Universal Robots URScript: test_4.script

def Machining2():
  # Default parameters:
  global speed_ms = 0.3
  global speed_rads = 0.75
  global accel_mss = 3
  global accel_radss = 1.2
  global blend_radius_m = 0.001

  # Add subprograms here
  # Start of main program
  # Program generated by RoboDK v5.6.5 for UR10e on 02/02/2024 11:53:03
  # Using nominal kinematics.
  blend_radius_m = 0.002
  speed_ms = 1.000
  # set_reference(p[0.335000, -0.152000, -0.013000, 0.000000, 0.000000, 0.000000])
  set_tcp(p[0.000000, 0.000000, 0.252000, 0.000000, 0.000000, 0.000000])
  # Show Tool
  movej([0.067194, -1.005485, -2.507684, -1.199220, 1.570796, 1.637990],accel_radss,speed_rads,0,blend_radius_m)
  movel([0.067194, -1.005485, -2.507684, -1.199220, 1.570796, 1.637990],accel_mss,speed_ms,0,blend_radius_m)
  # Splitting Linear movement in 6 (instruction 7: MoveL 3)
  movel([0.067194, -1.023371, -2.532341, -1.156677, 1.570796, 1.637990],accel_mss,speed_ms,0,blend_radius_m)
  movel([0.067194, -1.043822, -2.556463, -1.112104, 1.570796, 1.637990],accel_mss,speed_ms,0,blend_radius_m)
  movel([0.067194, -1.067076, -2.580006, -1.065307, 1.570796, 1.637990],accel_mss,speed_ms,0,blend_radius_m)
  movel([0.067194, -1.093389, -2.602916, -1.016084, 1.570796, 1.637990],accel_mss,speed_ms,0,blend_radius_m)
  movel([0.067194, -1.123035, -2.625130, -0.964224, 1.570796, 1.637990],accel_mss,speed_ms,0,blend_radius_m)
  movel([0.067194, -1.156300, -2.646577, -0.909512, 1.570796, 1.637990],accel_mss,speed_ms,0,blend_radius_m)
  movel([0.067194, -1.156300, -2.646577, -0.909512, 1.570796, 1.637990],accel_mss,speed_ms,0,blend_radius_m)
  speed_ms = 1.000
  movel([0.067194, -1.156300, -2.646577, -0.909512, 1.570796, 1.637990],accel_mss,speed_ms,0,blend_radius_m)
  movel([0.067194, -1.156300, -2.646577, -0.909512, 1.570796, 1.637990],accel_mss,speed_ms,0,blend_radius_m)
  movel([0.067194, -1.156300, -2.646577, -0.909512, 1.570796, 1.637990],accel_mss,speed_ms,0,blend_radius_m)
  speed_ms = 0.005
  # Splitting Linear movement in 2 (instruction 14: MoveL 8)
  movel([0.067194, -1.135891, -2.633806, -0.942693, 1.570796, 1.637990],accel_mss,speed_ms,0,blend_radius_m)
  movel([0.067194, -1.116825, -2.620746, -0.974817, 1.570796, 1.637990],accel_mss,speed_ms,0,blend_radius_m)
  speed_ms = 1.000
  # Splitting Linear movement in 2 (instruction 16: MoveL 9)
  movel([0.067194, -1.135891, -2.633806, -0.942693, 1.570796, 1.637990],accel_mss,speed_ms,0,blend_radius_m)
  movel([0.067194, -1.156300, -2.646577, -0.909512, 1.570796, 1.637990],accel_mss,speed_ms,0,blend_radius_m)
  speed_ms = 0.040
  movel([0.067194, -1.156300, -2.646577, -0.909512, 1.570796, 1.637990],accel_mss,speed_ms,0,blend_radius_m)
  speed_ms = 1.000
  movel([0.067194, -1.156300, -2.646577, -0.909512, 1.570796, 1.637990],accel_mss,speed_ms,0,blend_radius_m)
  # Splitting Linear movement in 8 (instruction 21: MoveL 12)
  movel([0.093765, -1.178967, -2.636050, -0.897372, 1.570796, 1.664562],accel_mss,speed_ms,0,blend_radius_m)
  movel([0.118639, -1.202315, -2.624642, -0.885432, 1.570796, 1.689436],accel_mss,speed_ms,0,blend_radius_m)
  movel([0.141916, -1.226161, -2.612379, -0.873849, 1.570796, 1.712712],accel_mss,speed_ms,0,blend_radius_m)
  movel([0.163698, -1.250347, -2.599285, -0.862758, 1.570796, 1.734494],accel_mss,speed_ms,0,blend_radius_m)
  movel([0.184083, -1.274733, -2.585389, -0.852267, 1.570796, 1.754880],accel_mss,speed_ms,0,blend_radius_m)
  movel([0.203170, -1.299204, -2.570720, -0.842465, 1.570796, 1.773967],accel_mss,speed_ms,0,blend_radius_m)
  movel([0.221051, -1.323665, -2.555309, -0.833415, 1.570796, 1.791848],accel_mss,speed_ms,0,blend_radius_m)
  movel([0.237813, -1.348037, -2.539186, -0.825166, 1.570796, 1.808610],accel_mss,speed_ms,0,blend_radius_m)
  speed_ms = 0.005
  movel([0.237813, -1.389023, -2.559646, -0.763720, 1.570796, 1.808610],accel_mss,speed_ms,0,blend_radius_m)
  speed_ms = 0.025
  movel([0.235045, -1.393576, -2.556354, -0.762459, 1.570796, 1.805842],accel_mss,speed_ms,0,blend_radius_m)
  movel([0.233553, -1.395826, -2.554716, -0.761847, 1.570796, 1.804349],accel_mss,speed_ms,0,blend_radius_m)
  movel([0.231969, -1.398040, -2.553098, -0.761252, 1.570796, 1.802766],accel_mss,speed_ms,0,blend_radius_m)
  movel([0.230284, -1.400201, -2.551510, -0.760677, 1.570796, 1.801081],accel_mss,speed_ms,0,blend_radius_m)
  movel([0.228485, -1.402296, -2.549965, -0.760127, 1.570796, 1.799282],accel_mss,speed_ms,0,blend_radius_m)
  movel([0.226558, -1.404312, -2.548473, -0.759604, 1.570796, 1.797355],accel_mss,speed_ms,0,blend_radius_m)
  movel([0.224490, -1.406231, -2.547046, -0.759112, 1.570796, 1.795286],accel_mss,speed_ms,0,blend_radius_m)
  movel([0.225289, -1.405338, -2.547711, -0.759341, 1.570796, 1.796085],accel_mss,speed_ms,0,blend_radius_m)
  movel([0.226090, -1.404119, -2.548616, -0.759654, 1.570796, 1.796886],accel_mss,speed_ms,0,blend_radius_m)
  movel([0.226657, -1.402885, -2.549530, -0.759974, 1.570796, 1.797453],accel_mss,speed_ms,0,blend_radius_m)
  movel([0.226775, -1.402364, -2.549915, -0.760110, 1.570796, 1.797572],accel_mss,speed_ms,0,blend_radius_m)
  movel([0.226747, -1.401956, -2.550216, -0.760216, 1.570796, 1.797543],accel_mss,speed_ms,0,blend_radius_m)
  movel([0.226540, -1.401693, -2.550411, -0.760285, 1.570796, 1.797336],accel_mss,speed_ms,0,blend_radius_m)
  movel([0.226190, -1.401646, -2.550445, -0.760297, 1.570796, 1.796986],accel_mss,speed_ms,0,blend_radius_m)
  movel([0.225721, -1.401788, -2.550341, -0.760260, 1.570796, 1.796518],accel_mss,speed_ms,0,blend_radius_m)
  movel([0.225147, -1.402096, -2.550113, -0.760180, 1.570796, 1.795944],accel_mss,speed_ms,0,blend_radius_m)
  movel([0.223775, -1.403102, -2.549370, -0.759918, 1.570796, 1.794571],accel_mss,speed_ms,0,blend_radius_m)
  movel([0.222231, -1.404457, -2.548365, -0.759567, 1.570796, 1.793027],accel_mss,speed_ms,0,blend_radius_m)
  movel([0.219245, -1.407409, -2.546167, -0.758812, 1.570796, 1.790041],accel_mss,speed_ms,0,blend_radius_m)
  movel([0.217410, -1.409332, -2.544729, -0.758328, 1.570796, 1.788207],accel_mss,speed_ms,0,blend_radius_m)
  movel([0.214705, -1.411968, -2.542749, -0.757672, 1.570796, 1.785501],accel_mss,speed_ms,0,blend_radius_m)
  movel([0.213250, -1.413159, -2.541851, -0.757379, 1.570796, 1.784046],accel_mss,speed_ms,0,blend_radius_m)
  movel([0.211689, -1.414182, -2.541078, -0.757129, 1.570796, 1.782486],accel_mss,speed_ms,0,blend_radius_m)
  movel([0.212040, -1.413816, -2.541354, -0.757218, 1.570796, 1.782836],accel_mss,speed_ms,0,blend_radius_m)
  movel([0.212351, -1.413193, -2.541825, -0.757371, 1.570796, 1.783147],accel_mss,speed_ms,0,blend_radius_m)
  movel([0.212822, -1.411511, -2.543093, -0.757785, 1.570796, 1.783618],accel_mss,speed_ms,0,blend_radius_m)
  movel([0.213027, -1.409824, -2.544360, -0.758204, 1.570796, 1.783823],accel_mss,speed_ms,0,blend_radius_m)
  movel([0.213004, -1.409193, -2.544834, -0.758363, 1.570796, 1.783800],accel_mss,speed_ms,0,blend_radius_m)
  movel([0.212886, -1.408822, -2.545111, -0.758456, 1.570796, 1.783683],accel_mss,speed_ms,0,blend_radius_m)
  movel([0.212415, -1.408436, -2.545400, -0.758553, 1.570796, 1.783211],accel_mss,speed_ms,0,blend_radius_m)
  movel([0.211885, -1.408340, -2.545472, -0.758577, 1.570796, 1.782681],accel_mss,speed_ms,0,blend_radius_m)
  movel([0.211310, -1.408476, -2.545370, -0.758543, 1.570796, 1.782107],accel_mss,speed_ms,0,blend_radius_m)
  movel([0.210707, -1.408794, -2.545132, -0.758463, 1.570796, 1.781503],accel_mss,speed_ms,0,blend_radius_m)
  movel([0.209488, -1.409732, -2.544429, -0.758227, 1.570796, 1.780285],accel_mss,speed_ms,0,blend_radius_m)
  movel([0.208361, -1.410705, -2.543699, -0.757985, 1.570796, 1.779157],accel_mss,speed_ms,0,blend_radius_m)
  movel([0.206539, -1.412115, -2.542638, -0.757636, 1.570796, 1.777335],accel_mss,speed_ms,0,blend_radius_m)
  movel([0.204719, -1.413331, -2.541721, -0.757337, 1.570796, 1.775515],accel_mss,speed_ms,0,blend_radius_m)
  movel([0.202815, -1.414308, -2.540982, -0.757099, 1.570796, 1.773611],accel_mss,speed_ms,0,blend_radius_m)
  movel([0.200751, -1.414992, -2.540465, -0.756933, 1.570796, 1.771548],accel_mss,speed_ms,0,blend_radius_m)
  movel([0.202050, -1.413855, -2.541325, -0.757209, 1.570796, 1.772846],accel_mss,speed_ms,0,blend_radius_m)
  movel([0.203160, -1.412607, -2.542267, -0.757515, 1.570796, 1.773956],accel_mss,speed_ms,0,blend_radius_m)
  movel([0.203562, -1.411917, -2.542787, -0.757685, 1.570796, 1.774359],accel_mss,speed_ms,0,blend_radius_m)
  movel([0.203796, -1.411225, -2.543308, -0.757856, 1.570796, 1.774592],accel_mss,speed_ms,0,blend_radius_m)
  movel([0.203827, -1.410587, -2.543788, -0.758014, 1.570796, 1.774624],accel_mss,speed_ms,0,blend_radius_m)
  movel([0.203610, -1.410065, -2.544180, -0.758144, 1.570796, 1.774406],accel_mss,speed_ms,0,blend_radius_m)
  movel([0.203000, -1.409678, -2.544470, -0.758241, 1.570796, 1.773797],accel_mss,speed_ms,0,blend_radius_m)
  movel([0.202157, -1.409585, -2.544540, -0.758264, 1.570796, 1.772954],accel_mss,speed_ms,0,blend_radius_m)
  movel([0.201181, -1.409700, -2.544453, -0.758235, 1.570796, 1.771977],accel_mss,speed_ms,0,blend_radius_m)
  movel([0.200179, -1.409929, -2.544282, -0.758178, 1.570796, 1.770975],accel_mss,speed_ms,0,blend_radius_m)
  speed_ms = 0.005
  movel([0.200179, -1.401572, -2.540395, -0.770422, 1.570796, 1.770975],accel_mss,speed_ms,0,blend_radius_m)
  speed_ms = 0.040
  movel([0.198845, -1.420778, -2.525900, -0.765711, 1.570796, 1.769641],accel_mss,speed_ms,0,blend_radius_m)
  speed_ms = 0.005
  movel([0.198845, -1.428998, -2.529707, -0.753685, 1.570796, 1.769641],accel_mss,speed_ms,0,blend_radius_m)
  speed_ms = 0.025
  movel([0.199509, -1.427856, -2.530594, -0.753939, 1.570796, 1.770306],accel_mss,speed_ms,0,blend_radius_m)
  movel([0.200309, -1.426742, -2.531459, -0.754188, 1.570796, 1.771105],accel_mss,speed_ms,0,blend_radius_m)
  movel([0.201225, -1.425672, -2.532287, -0.754429, 1.570796, 1.772021],accel_mss,speed_ms,0,blend_radius_m)
  movel([0.202246, -1.424659, -2.533070, -0.754660, 1.570796, 1.773042],accel_mss,speed_ms,0,blend_radius_m)
  movel([0.203354, -1.423716, -2.533798, -0.754875, 1.570796, 1.774151],accel_mss,speed_ms,0,blend_radius_m)
  movel([0.204537, -1.422860, -2.534457, -0.755072, 1.570796, 1.775333],accel_mss,speed_ms,0,blend_radius_m)
  movel([0.205775, -1.422105, -2.535038, -0.755247, 1.570796, 1.776572],accel_mss,speed_ms,0,blend_radius_m)
  movel([0.207059, -1.421462, -2.535531, -0.755396, 1.570796, 1.777855],accel_mss,speed_ms,0,blend_radius_m)
  movel([0.208994, -1.420727, -2.536094, -0.755567, 1.570796, 1.779790],accel_mss,speed_ms,0,blend_radius_m)
  movel([0.210833, -1.420284, -2.536434, -0.755671, 1.570796, 1.781629],accel_mss,speed_ms,0,blend_radius_m)
  movel([0.212575, -1.420109, -2.536568, -0.755712, 1.570796, 1.783371],accel_mss,speed_ms,0,blend_radius_m)
  movel([0.214215, -1.420179, -2.536514, -0.755696, 1.570796, 1.785012],accel_mss,speed_ms,0,blend_radius_m)
  movel([0.215754, -1.420471, -2.536291, -0.755627, 1.570796, 1.786550],accel_mss,speed_ms,0,blend_radius_m)
  movel([0.217191, -1.420963, -2.535914, -0.755512, 1.570796, 1.787988],accel_mss,speed_ms,0,blend_radius_m)
  movel([0.218522, -1.421632, -2.535400, -0.755356, 1.570796, 1.789319],accel_mss,speed_ms,0,blend_radius_m)
  movel([0.219749, -1.422454, -2.534769, -0.755166, 1.570796, 1.790545],accel_mss,speed_ms,0,blend_radius_m)
  movel([0.220869, -1.423406, -2.534037, -0.754946, 1.570796, 1.791665],accel_mss,speed_ms,0,blend_radius_m)
  movel([0.221883, -1.424465, -2.533220, -0.754704, 1.570796, 1.792680],accel_mss,speed_ms,0,blend_radius_m)
  movel([0.223597, -1.426808, -2.531407, -0.754173, 1.570796, 1.794393],accel_mss,speed_ms,0,blend_radius_m)
  movel([0.224891, -1.429295, -2.529475, -0.753619, 1.570796, 1.795688],accel_mss,speed_ms,0,blend_radius_m)
  movel([0.225764, -1.431748, -2.527560, -0.753082, 1.570796, 1.796561],accel_mss,speed_ms,0,blend_radius_m)
  movel([0.226370, -1.434419, -2.525463, -0.752506, 1.570796, 1.797167],accel_mss,speed_ms,0,blend_radius_m)
  movel([0.226742, -1.437185, -2.523282, -0.751922, 1.570796, 1.797539],accel_mss,speed_ms,0,blend_radius_m)
  movel([0.226909, -1.440026, -2.521029, -0.751334, 1.570796, 1.797705],accel_mss,speed_ms,0,blend_radius_m)
  movel([0.226896, -1.442925, -2.518717, -0.750747, 1.570796, 1.797692],accel_mss,speed_ms,0,blend_radius_m)
  movel([0.226731, -1.445864, -2.516361, -0.750164, 1.570796, 1.797527],accel_mss,speed_ms,0,blend_radius_m)
  movel([0.226444, -1.448825, -2.513973, -0.749591, 1.570796, 1.797240],accel_mss,speed_ms,0,blend_radius_m)
  movel([0.225607, -1.454748, -2.509158, -0.748483, 1.570796, 1.796403],accel_mss,speed_ms,0,blend_radius_m)
  movel([0.224989, -1.458871, -2.505774, -0.747744, 1.570796, 1.795785],accel_mss,speed_ms,0,blend_radius_m)
  movel([0.224859, -1.460871, -2.504123, -0.747395, 1.570796, 1.795655],accel_mss,speed_ms,0,blend_radius_m)
  movel([0.224966, -1.462787, -2.502536, -0.747066, 1.570796, 1.795762],accel_mss,speed_ms,0,blend_radius_m)
  movel([0.225466, -1.465173, -2.500551, -0.746665, 1.570796, 1.796262],accel_mss,speed_ms,0,blend_radius_m)
  movel([0.225968, -1.467564, -2.498554, -0.746271, 1.570796, 1.796765],accel_mss,speed_ms,0,blend_radius_m)
  movel([0.226065, -1.468777, -2.497537, -0.746075, 1.570796, 1.796861],accel_mss,speed_ms,0,blend_radius_m)
  movel([0.225974, -1.470011, -2.496500, -0.745878, 1.570796, 1.796771],accel_mss,speed_ms,0,blend_radius_m)
  movel([0.225636, -1.471270, -2.495440, -0.745679, 1.570796, 1.796433],accel_mss,speed_ms,0,blend_radius_m)
  movel([0.224991, -1.472564, -2.494348, -0.745477, 1.570796, 1.795787],accel_mss,speed_ms,0,blend_radius_m)
  movel([0.226901, -1.469422, -2.496996, -0.745972, 1.570796, 1.797697],accel_mss,speed_ms,0,blend_radius_m)
  movel([0.228644, -1.466259, -2.499645, -0.746485, 1.570796, 1.799440],accel_mss,speed_ms,0,blend_radius_m)
  movel([0.231835, -1.459849, -2.504967, -0.747573, 1.570796, 1.802632],accel_mss,speed_ms,0,blend_radius_m)
  movel([0.233501, -1.456244, -2.507933, -0.748212, 1.570796, 1.804297],accel_mss,speed_ms,0,blend_radius_m)
  movel([0.235068, -1.452620, -2.510894, -0.748875, 1.570796, 1.805865],accel_mss,speed_ms,0,blend_radius_m)
  movel([0.237984, -1.445308, -2.516808, -0.750274, 1.570796, 1.808780],accel_mss,speed_ms,0,blend_radius_m)
  movel([0.240604, -1.438082, -2.522572, -0.751735, 1.570796, 1.811400],accel_mss,speed_ms,0,blend_radius_m)
  movel([0.241738, -1.434441, -2.525447, -0.752502, 1.570796, 1.812534],accel_mss,speed_ms,0,blend_radius_m)
  movel([0.242662, -1.430833, -2.528275, -0.753281, 1.570796, 1.813459],accel_mss,speed_ms,0,blend_radius_m)
  movel([0.243176, -1.428019, -2.530468, -0.753902, 1.570796, 1.813972],accel_mss,speed_ms,0,blend_radius_m)
  movel([0.243556, -1.425209, -2.532645, -0.754534, 1.570796, 1.814353],accel_mss,speed_ms,0,blend_radius_m)
  movel([0.243953, -1.422370, -2.534833, -0.755185, 1.570796, 1.814749],accel_mss,speed_ms,0,blend_radius_m)
  movel([0.244515, -1.419469, -2.537057, -0.755863, 1.570796, 1.815311],accel_mss,speed_ms,0,blend_radius_m)
  movel([0.244763, -1.418683, -2.537657, -0.756048, 1.570796, 1.815560],accel_mss,speed_ms,0,blend_radius_m)
  movel([0.245167, -1.417894, -2.538259, -0.756236, 1.570796, 1.815963],accel_mss,speed_ms,0,blend_radius_m)
  movel([0.245733, -1.417238, -2.538759, -0.756392, 1.570796, 1.816529],accel_mss,speed_ms,0,blend_radius_m)
  movel([0.246084, -1.417001, -2.538939, -0.756449, 1.570796, 1.816880],accel_mss,speed_ms,0,blend_radius_m)
  movel([0.246482, -1.416844, -2.539058, -0.756486, 1.570796, 1.817278],accel_mss,speed_ms,0,blend_radius_m)
  movel([0.247021, -1.416802, -2.539091, -0.756496, 1.570796, 1.817817],accel_mss,speed_ms,0,blend_radius_m)
  movel([0.247506, -1.416887, -2.539026, -0.756476, 1.570796, 1.818302],accel_mss,speed_ms,0,blend_radius_m)
  movel([0.249997, -1.417659, -2.538438, -0.756291, 1.570796, 1.820793],accel_mss,speed_ms,0,blend_radius_m)
  movel([0.252171, -1.418695, -2.537648, -0.756045, 1.570796, 1.822967],accel_mss,speed_ms,0,blend_radius_m)
  movel([0.254051, -1.419966, -2.536677, -0.755746, 1.570796, 1.824848],accel_mss,speed_ms,0,blend_radius_m)
  movel([0.255662, -1.421454, -2.535537, -0.755398, 1.570796, 1.826458],accel_mss,speed_ms,0,blend_radius_m)
  movel([0.257025, -1.423131, -2.534248, -0.755010, 1.570796, 1.827822],accel_mss,speed_ms,0,blend_radius_m)
  movel([0.258167, -1.424975, -2.532827, -0.754588, 1.570796, 1.828963],accel_mss,speed_ms,0,blend_radius_m)
  movel([0.259109, -1.426961, -2.531289, -0.754139, 1.570796, 1.829905],accel_mss,speed_ms,0,blend_radius_m)
  movel([0.259873, -1.429069, -2.529651, -0.753669, 1.570796, 1.830669],accel_mss,speed_ms,0,blend_radius_m)
  movel([0.260485, -1.431275, -2.527930, -0.753184, 1.570796, 1.831281],accel_mss,speed_ms,0,blend_radius_m)
  movel([0.260970, -1.433556, -2.526142, -0.752691, 1.570796, 1.831766],accel_mss,speed_ms,0,blend_radius_m)
  movel([0.261645, -1.438257, -2.522433, -0.751699, 1.570796, 1.832442],accel_mss,speed_ms,0,blend_radius_m)
  movel([0.262466, -1.447636, -2.514933, -0.749819, 1.570796, 1.833262],accel_mss,speed_ms,0,blend_radius_m)
  movel([0.262681, -1.449067, -2.513777, -0.749544, 1.570796, 1.833478],accel_mss,speed_ms,0,blend_radius_m)
  movel([0.262929, -1.449701, -2.513264, -0.749424, 1.570796, 1.833725],accel_mss,speed_ms,0,blend_radius_m)
  movel([0.263331, -1.450229, -2.512836, -0.749323, 1.570796, 1.834127],accel_mss,speed_ms,0,blend_radius_m)
  movel([0.264227, -1.450735, -2.512426, -0.749228, 1.570796, 1.835023],accel_mss,speed_ms,0,blend_radius_m)
  movel([0.264740, -1.450835, -2.512345, -0.749209, 1.570796, 1.835536],accel_mss,speed_ms,0,blend_radius_m)
  movel([0.265289, -1.450841, -2.512340, -0.749208, 1.570796, 1.836086],accel_mss,speed_ms,0,blend_radius_m)
  movel([0.266462, -1.450615, -2.512524, -0.749250, 1.570796, 1.837259],accel_mss,speed_ms,0,blend_radius_m)
  movel([0.267692, -1.450120, -2.512925, -0.749344, 1.570796, 1.838488],accel_mss,speed_ms,0,blend_radius_m)
  movel([0.268921, -1.449427, -2.513487, -0.749476, 1.570796, 1.839717],accel_mss,speed_ms,0,blend_radius_m)
  movel([0.270093, -1.448599, -2.514156, -0.749634, 1.570796, 1.840889],accel_mss,speed_ms,0,blend_radius_m)
  movel([0.271154, -1.447703, -2.514880, -0.749807, 1.570796, 1.841950],accel_mss,speed_ms,0,blend_radius_m)
  movel([0.272041, -1.446803, -2.515605, -0.749981, 1.570796, 1.842837],accel_mss,speed_ms,0,blend_radius_m)
  movel([0.273423, -1.445193, -2.516900, -0.750296, 1.570796, 1.844219],accel_mss,speed_ms,0,blend_radius_m)
  movel([0.274736, -1.443535, -2.518229, -0.750625, 1.570796, 1.845533],accel_mss,speed_ms,0,blend_radius_m)
  movel([0.277146, -1.440108, -2.520963, -0.751317, 1.570796, 1.847942],accel_mss,speed_ms,0,blend_radius_m)
  movel([0.279260, -1.436587, -2.523754, -0.752048, 1.570796, 1.850057],accel_mss,speed_ms,0,blend_radius_m)
  movel([0.281063, -1.433036, -2.526550, -0.752803, 1.570796, 1.851859],accel_mss,speed_ms,0,blend_radius_m)
  movel([0.281687, -1.431692, -2.527603, -0.753094, 1.570796, 1.852483],accel_mss,speed_ms,0,blend_radius_m)
  movel([0.282425, -1.430374, -2.528634, -0.753382, 1.570796, 1.853221],accel_mss,speed_ms,0,blend_radius_m)
  movel([0.282883, -1.429754, -2.529117, -0.753518, 1.570796, 1.853679],accel_mss,speed_ms,0,blend_radius_m)
  movel([0.283426, -1.429173, -2.529570, -0.753646, 1.570796, 1.854222],accel_mss,speed_ms,0,blend_radius_m)
  movel([0.284071, -1.428643, -2.529982, -0.753763, 1.570796, 1.854867],accel_mss,speed_ms,0,blend_radius_m)
  movel([0.284836, -1.428179, -2.530343, -0.753867, 1.570796, 1.855633],accel_mss,speed_ms,0,blend_radius_m)
  movel([0.285921, -1.427810, -2.530630, -0.753949, 1.570796, 1.856718],accel_mss,speed_ms,0,blend_radius_m)
  movel([0.286948, -1.427790, -2.530645, -0.753953, 1.570796, 1.857744],accel_mss,speed_ms,0,blend_radius_m)
  movel([0.287857, -1.428051, -2.530443, -0.753895, 1.570796, 1.858653],accel_mss,speed_ms,0,blend_radius_m)
  movel([0.288594, -1.428522, -2.530077, -0.753790, 1.570796, 1.859391],accel_mss,speed_ms,0,blend_radius_m)
  movel([0.289573, -1.429534, -2.529289, -0.753566, 1.570796, 1.860369],accel_mss,speed_ms,0,blend_radius_m)
  movel([0.290398, -1.430690, -2.528386, -0.753312, 1.570796, 1.861194],accel_mss,speed_ms,0,blend_radius_m)
  movel([0.291712, -1.433202, -2.526420, -0.752767, 1.570796, 1.862509],accel_mss,speed_ms,0,blend_radius_m)
  movel([0.292196, -1.434457, -2.525434, -0.752498, 1.570796, 1.862993],accel_mss,speed_ms,0,blend_radius_m)
  movel([0.292534, -1.435746, -2.524418, -0.752225, 1.570796, 1.863331],accel_mss,speed_ms,0,blend_radius_m)
  movel([0.292737, -1.437066, -2.523376, -0.751947, 1.570796, 1.863533],accel_mss,speed_ms,0,blend_radius_m)
  movel([0.292810, -1.438415, -2.522308, -0.751666, 1.570796, 1.863606],accel_mss,speed_ms,0,blend_radius_m)
  movel([0.292761, -1.439788, -2.521218, -0.751383, 1.570796, 1.863557],accel_mss,speed_ms,0,blend_radius_m)
  movel([0.292327, -1.442600, -2.518977, -0.750812, 1.570796, 1.863123],accel_mss,speed_ms,0,blend_radius_m)
  movel([0.291955, -1.444032, -2.517831, -0.750526, 1.570796, 1.862752],accel_mss,speed_ms,0,blend_radius_m)
  movel([0.290947, -1.446934, -2.515500, -0.749956, 1.570796, 1.861744],accel_mss,speed_ms,0,blend_radius_m)
  movel([0.289630, -1.449867, -2.513130, -0.749392, 1.570796, 1.860426],accel_mss,speed_ms,0,blend_radius_m)
  movel([0.288058, -1.452813, -2.510736, -0.748839, 1.570796, 1.858855],accel_mss,speed_ms,0,blend_radius_m)
  movel([0.286295, -1.455747, -2.508340, -0.748302, 1.570796, 1.857091],accel_mss,speed_ms,0,blend_radius_m)
  movel([0.283469, -1.459970, -2.504868, -0.747552, 1.570796, 1.854265],accel_mss,speed_ms,0,blend_radius_m)
  movel([0.281933, -1.462043, -2.503153, -0.747193, 1.570796, 1.852729],accel_mss,speed_ms,0,blend_radius_m)
  movel([0.280302, -1.464070, -2.501470, -0.746849, 1.570796, 1.851098],accel_mss,speed_ms,0,blend_radius_m)
  movel([0.278570, -1.466034, -2.499833, -0.746522, 1.570796, 1.849366],accel_mss,speed_ms,0,blend_radius_m)
  movel([0.276731, -1.467921, -2.498255, -0.746213, 1.570796, 1.847527],accel_mss,speed_ms,0,blend_radius_m)
  movel([0.274770, -1.469718, -2.496747, -0.745924, 1.570796, 1.845566],accel_mss,speed_ms,0,blend_radius_m)
  movel([0.272685, -1.471406, -2.495325, -0.745657, 1.570796, 1.843481],accel_mss,speed_ms,0,blend_radius_m)
  movel([0.269604, -1.473590, -2.493480, -0.745319, 1.570796, 1.840400],accel_mss,speed_ms,0,blend_radius_m)
  movel([0.267919, -1.474637, -2.492594, -0.745159, 1.570796, 1.838716],accel_mss,speed_ms,0,blend_radius_m)
  movel([0.266184, -1.475578, -2.491795, -0.745017, 1.570796, 1.836981],accel_mss,speed_ms,0,blend_radius_m)
  movel([0.264435, -1.476358, -2.491131, -0.744900, 1.570796, 1.835232],accel_mss,speed_ms,0,blend_radius_m)
  movel([0.262707, -1.476922, -2.490651, -0.744816, 1.570796, 1.833504],accel_mss,speed_ms,0,blend_radius_m)
  movel([0.261035, -1.477213, -2.490403, -0.744773, 1.570796, 1.831831],accel_mss,speed_ms,0,blend_radius_m)
  movel([0.260230, -1.477239, -2.490381, -0.744769, 1.570796, 1.831026],accel_mss,speed_ms,0,blend_radius_m)
  movel([0.259454, -1.477175, -2.490436, -0.744778, 1.570796, 1.830251],accel_mss,speed_ms,0,blend_radius_m)
  movel([0.258632, -1.476991, -2.490592, -0.744806, 1.570796, 1.829428],accel_mss,speed_ms,0,blend_radius_m)
  movel([0.257902, -1.476699, -2.490841, -0.744849, 1.570796, 1.828698],accel_mss,speed_ms,0,blend_radius_m)
  movel([0.257255, -1.476309, -2.491173, -0.744907, 1.570796, 1.828051],accel_mss,speed_ms,0,blend_radius_m)
  movel([0.256688, -1.475830, -2.491580, -0.744979, 1.570796, 1.827484],accel_mss,speed_ms,0,blend_radius_m)
  movel([0.255764, -1.474653, -2.492580, -0.745156, 1.570796, 1.826560],accel_mss,speed_ms,0,blend_radius_m)
  movel([0.255085, -1.473246, -2.493771, -0.745371, 1.570796, 1.825882],accel_mss,speed_ms,0,blend_radius_m)
  movel([0.254602, -1.471698, -2.495080, -0.745612, 1.570796, 1.825398],accel_mss,speed_ms,0,blend_radius_m)
  movel([0.254267, -1.470090, -2.496434, -0.745865, 1.570796, 1.825064],accel_mss,speed_ms,0,blend_radius_m)
  movel([0.253855, -1.467040, -2.498992, -0.746357, 1.570796, 1.824652],accel_mss,speed_ms,0,blend_radius_m)
  movel([0.253682, -1.465611, -2.500186, -0.746592, 1.570796, 1.824478],accel_mss,speed_ms,0,blend_radius_m)
  movel([0.253352, -1.464264, -2.501308, -0.746817, 1.570796, 1.824148],accel_mss,speed_ms,0,blend_radius_m)
  movel([0.253057, -1.463681, -2.501793, -0.746915, 1.570796, 1.823853],accel_mss,speed_ms,0,blend_radius_m)
  movel([0.252636, -1.463189, -2.502202, -0.746998, 1.570796, 1.823432],accel_mss,speed_ms,0,blend_radius_m)
  movel([0.252062, -1.462813, -2.502514, -0.747062, 1.570796, 1.822858],accel_mss,speed_ms,0,blend_radius_m)
  movel([0.251306, -1.462576, -2.502711, -0.747102, 1.570796, 1.822103],accel_mss,speed_ms,0,blend_radius_m)
  movel([0.251464, -1.462664, -2.502638, -0.747087, 1.570796, 1.822260],accel_mss,speed_ms,0,blend_radius_m)
  movel([0.251531, -1.462846, -2.502487, -0.747056, 1.570796, 1.822327],accel_mss,speed_ms,0,blend_radius_m)
  movel([0.251409, -1.463470, -2.501968, -0.746950, 1.570796, 1.822205],accel_mss,speed_ms,0,blend_radius_m)
  movel([0.250980, -1.464398, -2.501197, -0.746794, 1.570796, 1.821777],accel_mss,speed_ms,0,blend_radius_m)
  movel([0.250294, -1.465582, -2.500210, -0.746597, 1.570796, 1.821091],accel_mss,speed_ms,0,blend_radius_m)
  movel([0.248323, -1.468516, -2.497756, -0.746117, 1.570796, 1.819119],accel_mss,speed_ms,0,blend_radius_m)
  movel([0.245847, -1.471879, -2.494927, -0.745583, 1.570796, 1.816643],accel_mss,speed_ms,0,blend_radius_m)
  movel([0.240761, -1.478352, -2.489431, -0.744605, 1.570796, 1.811557],accel_mss,speed_ms,0,blend_radius_m)
  movel([0.237727, -1.481981, -2.486322, -0.744086, 1.570796, 1.808524],accel_mss,speed_ms,0,blend_radius_m)
  movel([0.234260, -1.485603, -2.483198, -0.743587, 1.570796, 1.805057],accel_mss,speed_ms,0,blend_radius_m)
  movel([0.230760, -1.489122, -2.480145, -0.743123, 1.570796, 1.801556],accel_mss,speed_ms,0,blend_radius_m)
  movel([0.227207, -1.492577, -2.477127, -0.742685, 1.570796, 1.798003],accel_mss,speed_ms,0,blend_radius_m)
  movel([0.220164, -1.499147, -2.471337, -0.741905, 1.570796, 1.790960],accel_mss,speed_ms,0,blend_radius_m)
  movel([0.216634, -1.502153, -2.468665, -0.741571, 1.570796, 1.787430],accel_mss,speed_ms,0,blend_radius_m)
  movel([0.214805, -1.503553, -2.467416, -0.741420, 1.570796, 1.785601],accel_mss,speed_ms,0,blend_radius_m)
  movel([0.212926, -1.504857, -2.466250, -0.741282, 1.570796, 1.783722],accel_mss,speed_ms,0,blend_radius_m)
  movel([0.210985, -1.506044, -2.465186, -0.741159, 1.570796, 1.781781],accel_mss,speed_ms,0,blend_radius_m)
  movel([0.208979, -1.507094, -2.464243, -0.741052, 1.570796, 1.779776],accel_mss,speed_ms,0,blend_radius_m)
  movel([0.209952, -1.503854, -2.467147, -0.741388, 1.570796, 1.780748],accel_mss,speed_ms,0,blend_radius_m)
  movel([0.210102, -1.502910, -2.467991, -0.741489, 1.570796, 1.780898],accel_mss,speed_ms,0,blend_radius_m)
  movel([0.209998, -1.502528, -2.468331, -0.741530, 1.570796, 1.780794],accel_mss,speed_ms,0,blend_radius_m)
  movel([0.209695, -1.502293, -2.468540, -0.741555, 1.570796, 1.780492],accel_mss,speed_ms,0,blend_radius_m)
  movel([0.209319, -1.502260, -2.468570, -0.741559, 1.570796, 1.780116],accel_mss,speed_ms,0,blend_radius_m)
  movel([0.208897, -1.502355, -2.468485, -0.741549, 1.570796, 1.779693],accel_mss,speed_ms,0,blend_radius_m)
  movel([0.206817, -1.503186, -2.467744, -0.741459, 1.570796, 1.777613],accel_mss,speed_ms,0,blend_radius_m)
  movel([0.205619, -1.503492, -2.467471, -0.741426, 1.570796, 1.776415],accel_mss,speed_ms,0,blend_radius_m)
  movel([0.204447, -1.503636, -2.467342, -0.741411, 1.570796, 1.775243],accel_mss,speed_ms,0,blend_radius_m)
  movel([0.203332, -1.503615, -2.467361, -0.741413, 1.570796, 1.774128],accel_mss,speed_ms,0,blend_radius_m)
  movel([0.203014, -1.503515, -2.467451, -0.741424, 1.570796, 1.773811],accel_mss,speed_ms,0,blend_radius_m)
  movel([0.202959, -1.503290, -2.467651, -0.741448, 1.570796, 1.773755],accel_mss,speed_ms,0,blend_radius_m)
  movel([0.203433, -1.502377, -2.468465, -0.741546, 1.570796, 1.774229],accel_mss,speed_ms,0,blend_radius_m)
  movel([0.203455, -1.502071, -2.468738, -0.741580, 1.570796, 1.774251],accel_mss,speed_ms,0,blend_radius_m)
  movel([0.203315, -1.501832, -2.468951, -0.741606, 1.570796, 1.774111],accel_mss,speed_ms,0,blend_radius_m)
  movel([0.203056, -1.501676, -2.469090, -0.741623, 1.570796, 1.773853],accel_mss,speed_ms,0,blend_radius_m)
  movel([0.202724, -1.501620, -2.469140, -0.741629, 1.570796, 1.773520],accel_mss,speed_ms,0,blend_radius_m)
  movel([0.201977, -1.501757, -2.469018, -0.741614, 1.570796, 1.772773],accel_mss,speed_ms,0,blend_radius_m)
  movel([0.196468, -1.504100, -2.466928, -0.741362, 1.570796, 1.767264],accel_mss,speed_ms,0,blend_radius_m)
  movel([0.198143, -1.503132, -2.467792, -0.741465, 1.570796, 1.768940],accel_mss,speed_ms,0,blend_radius_m)
  movel([0.199814, -1.502046, -2.468761, -0.741582, 1.570796, 1.770610],accel_mss,speed_ms,0,blend_radius_m)
  movel([0.201463, -1.500866, -2.469811, -0.741712, 1.570796, 1.772259],accel_mss,speed_ms,0,blend_radius_m)
  movel([0.203082, -1.499608, -2.470928, -0.741853, 1.570796, 1.773878],accel_mss,speed_ms,0,blend_radius_m)
  movel([0.206181, -1.496938, -2.473291, -0.742160, 1.570796, 1.776977],accel_mss,speed_ms,0,blend_radius_m)
  movel([0.209010, -1.494195, -2.475707, -0.742487, 1.570796, 1.779806],accel_mss,speed_ms,0,blend_radius_m)
  movel([0.211927, -1.491138, -2.478386, -0.742865, 1.570796, 1.782723],accel_mss,speed_ms,0,blend_radius_m)
  movel([0.214736, -1.487976, -2.481141, -0.743272, 1.570796, 1.785533],accel_mss,speed_ms,0,blend_radius_m)
  movel([0.216063, -1.486353, -2.482549, -0.743487, 1.570796, 1.786859],accel_mss,speed_ms,0,blend_radius_m)
  movel([0.217321, -1.484701, -2.483978, -0.743709, 1.570796, 1.788118],accel_mss,speed_ms,0,blend_radius_m)
  movel([0.218492, -1.483021, -2.485427, -0.743940, 1.570796, 1.789289],accel_mss,speed_ms,0,blend_radius_m)
  movel([0.219565, -1.481308, -2.486900, -0.744180, 1.570796, 1.790361],accel_mss,speed_ms,0,blend_radius_m)
  movel([0.220151, -1.480225, -2.487830, -0.744335, 1.570796, 1.790948],accel_mss,speed_ms,0,blend_radius_m)
  movel([0.220648, -1.479122, -2.488774, -0.744493, 1.570796, 1.791444],accel_mss,speed_ms,0,blend_radius_m)
  movel([0.221390, -1.476879, -2.490688, -0.744822, 1.570796, 1.792187],accel_mss,speed_ms,0,blend_radius_m)
  movel([0.221820, -1.474621, -2.492607, -0.745161, 1.570796, 1.792616],accel_mss,speed_ms,0,blend_radius_m)
  movel([0.221961, -1.472385, -2.494499, -0.745505, 1.570796, 1.792757],accel_mss,speed_ms,0,blend_radius_m)
  movel([0.221848, -1.470210, -2.496333, -0.745846, 1.570796, 1.792644],accel_mss,speed_ms,0,blend_radius_m)
  movel([0.221510, -1.468134, -2.498076, -0.746179, 1.570796, 1.792307],accel_mss,speed_ms,0,blend_radius_m)
  movel([0.220973, -1.466199, -2.499695, -0.746495, 1.570796, 1.791770],accel_mss,speed_ms,0,blend_radius_m)
  movel([0.220271, -1.464442, -2.501160, -0.746787, 1.570796, 1.791067],accel_mss,speed_ms,0,blend_radius_m)
  movel([0.219658, -1.463586, -2.501872, -0.746931, 1.570796, 1.790454],accel_mss,speed_ms,0,blend_radius_m)
  movel([0.218810, -1.463040, -2.502325, -0.747023, 1.570796, 1.789606],accel_mss,speed_ms,0,blend_radius_m)
  movel([0.217785, -1.462799, -2.502526, -0.747064, 1.570796, 1.788581],accel_mss,speed_ms,0,blend_radius_m)
  movel([0.216644, -1.462855, -2.502480, -0.747055, 1.570796, 1.787440],accel_mss,speed_ms,0,blend_radius_m)
  movel([0.215441, -1.463197, -2.502196, -0.746997, 1.570796, 1.786237],accel_mss,speed_ms,0,blend_radius_m)
  movel([0.214235, -1.463817, -2.501680, -0.746892, 1.570796, 1.785031],accel_mss,speed_ms,0,blend_radius_m)
  movel([0.213088, -1.464705, -2.500941, -0.746743, 1.570796, 1.783884],accel_mss,speed_ms,0,blend_radius_m)
  movel([0.212056, -1.465849, -2.499987, -0.746553, 1.570796, 1.782852],accel_mss,speed_ms,0,blend_radius_m)
  movel([0.210631, -1.467673, -2.498463, -0.746254, 1.570796, 1.781428],accel_mss,speed_ms,0,blend_radius_m)
  movel([0.209126, -1.469445, -2.496977, -0.745968, 1.570796, 1.779922],accel_mss,speed_ms,0,blend_radius_m)
  movel([0.207533, -1.471141, -2.495549, -0.745699, 1.570796, 1.778330],accel_mss,speed_ms,0,blend_radius_m)
  movel([0.205841, -1.472744, -2.494196, -0.745449, 1.570796, 1.776637],accel_mss,speed_ms,0,blend_radius_m)
  movel([0.204046, -1.474228, -2.492940, -0.745221, 1.570796, 1.774842],accel_mss,speed_ms,0,blend_radius_m)
  movel([0.202135, -1.475576, -2.491796, -0.745017, 1.570796, 1.772932],accel_mss,speed_ms,0,blend_radius_m)
  movel([0.200101, -1.476767, -2.490783, -0.744839, 1.570796, 1.770898],accel_mss,speed_ms,0,blend_radius_m)
  movel([0.197938, -1.477780, -2.489920, -0.744689, 1.570796, 1.768734],accel_mss,speed_ms,0,blend_radius_m)
  movel([0.196789, -1.478175, -2.489582, -0.744631, 1.570796, 1.767585],accel_mss,speed_ms,0,blend_radius_m)
  movel([0.195645, -1.478439, -2.489357, -0.744593, 1.570796, 1.766441],accel_mss,speed_ms,0,blend_radius_m)
  movel([0.193385, -1.478731, -2.489107, -0.744550, 1.570796, 1.764182],accel_mss,speed_ms,0,blend_radius_m)
  movel([0.191654, -1.478794, -2.489054, -0.744541, 1.570796, 1.762450],accel_mss,speed_ms,0,blend_radius_m)
  movel([0.190052, -1.478647, -2.489179, -0.744562, 1.570796, 1.760849],accel_mss,speed_ms,0,blend_radius_m)
  movel([0.188577, -1.478308, -2.489469, -0.744612, 1.570796, 1.759374],accel_mss,speed_ms,0,blend_radius_m)
  movel([0.187221, -1.477794, -2.489908, -0.744687, 1.570796, 1.758017],accel_mss,speed_ms,0,blend_radius_m)
  movel([0.185975, -1.477124, -2.490479, -0.744786, 1.570796, 1.756772],accel_mss,speed_ms,0,blend_radius_m)
  movel([0.184836, -1.476313, -2.491170, -0.744907, 1.570796, 1.755632],accel_mss,speed_ms,0,blend_radius_m)
  movel([0.183800, -1.475377, -2.491965, -0.745047, 1.570796, 1.754597],accel_mss,speed_ms,0,blend_radius_m)
  movel([0.182860, -1.474336, -2.492848, -0.745204, 1.570796, 1.753657],accel_mss,speed_ms,0,blend_radius_m)
  movel([0.182010, -1.473207, -2.493804, -0.745377, 1.570796, 1.752807],accel_mss,speed_ms,0,blend_radius_m)
  movel([0.181248, -1.472003, -2.494822, -0.745564, 1.570796, 1.752044],accel_mss,speed_ms,0,blend_radius_m)
  movel([0.179959, -1.469452, -2.496970, -0.745967, 1.570796, 1.750756],accel_mss,speed_ms,0,blend_radius_m)
  movel([0.178954, -1.466817, -2.499178, -0.746393, 1.570796, 1.749750],accel_mss,speed_ms,0,blend_radius_m)
  movel([0.178191, -1.464244, -2.501325, -0.746820, 1.570796, 1.748988],accel_mss,speed_ms,0,blend_radius_m)
  movel([0.177732, -1.462222, -2.503005, -0.747163, 1.570796, 1.748528],accel_mss,speed_ms,0,blend_radius_m)
  movel([0.177384, -1.460085, -2.504773, -0.747532, 1.570796, 1.748181],accel_mss,speed_ms,0,blend_radius_m)
  movel([0.177159, -1.457845, -2.506619, -0.747926, 1.570796, 1.747955],accel_mss,speed_ms,0,blend_radius_m)
  movel([0.177072, -1.455518, -2.508528, -0.748343, 1.570796, 1.747868],accel_mss,speed_ms,0,blend_radius_m)
  movel([0.177130, -1.453118, -2.510489, -0.748783, 1.570796, 1.747926],accel_mss,speed_ms,0,blend_radius_m)
  movel([0.177349, -1.450659, -2.512488, -0.749242, 1.570796, 1.748145],accel_mss,speed_ms,0,blend_radius_m)
  movel([0.177742, -1.448157, -2.514513, -0.749719, 1.570796, 1.748539],accel_mss,speed_ms,0,blend_radius_m)
  movel([0.178321, -1.445626, -2.516552, -0.750211, 1.570796, 1.749118],accel_mss,speed_ms,0,blend_radius_m)
  movel([0.179099, -1.443080, -2.518594, -0.750716, 1.570796, 1.749895],accel_mss,speed_ms,0,blend_radius_m)
  movel([0.180086, -1.440538, -2.520622, -0.751230, 1.570796, 1.750883],accel_mss,speed_ms,0,blend_radius_m)
  movel([0.181298, -1.438011, -2.522628, -0.751750, 1.570796, 1.752094],accel_mss,speed_ms,0,blend_radius_m)
  movel([0.182748, -1.435518, -2.524598, -0.752273, 1.570796, 1.753544],accel_mss,speed_ms,0,blend_radius_m)
  movel([0.184446, -1.433076, -2.526519, -0.752794, 1.570796, 1.755242],accel_mss,speed_ms,0,blend_radius_m)
  movel([0.186408, -1.430699, -2.528380, -0.753310, 1.570796, 1.757205],accel_mss,speed_ms,0,blend_radius_m)
  movel([0.188643, -1.428409, -2.530164, -0.753815, 1.570796, 1.759439],accel_mss,speed_ms,0,blend_radius_m)
  movel([0.191163, -1.426223, -2.531861, -0.754305, 1.570796, 1.761960],accel_mss,speed_ms,0,blend_radius_m)
  movel([0.192220, -1.425458, -2.532453, -0.754478, 1.570796, 1.763017],accel_mss,speed_ms,0,blend_radius_m)
  movel([0.192778, -1.425155, -2.532687, -0.754547, 1.570796, 1.763574],accel_mss,speed_ms,0,blend_radius_m)
  movel([0.193347, -1.424951, -2.532845, -0.754593, 1.570796, 1.764143],accel_mss,speed_ms,0,blend_radius_m)
  movel([0.194154, -1.424899, -2.532885, -0.754605, 1.570796, 1.764950],accel_mss,speed_ms,0,blend_radius_m)
  movel([0.194819, -1.425121, -2.532713, -0.754554, 1.570796, 1.765615],accel_mss,speed_ms,0,blend_radius_m)
  movel([0.195329, -1.425551, -2.532381, -0.754457, 1.570796, 1.766125],accel_mss,speed_ms,0,blend_radius_m)
  movel([0.195667, -1.426118, -2.531942, -0.754329, 1.570796, 1.766463],accel_mss,speed_ms,0,blend_radius_m)
  movel([0.196015, -1.427586, -2.530804, -0.753999, 1.570796, 1.766812],accel_mss,speed_ms,0,blend_radius_m)
  movel([0.196048, -1.429207, -2.529543, -0.753638, 1.570796, 1.766844],accel_mss,speed_ms,0,blend_radius_m)
  movel([0.195783, -1.432540, -2.526939, -0.752910, 1.570796, 1.766580],accel_mss,speed_ms,0,blend_radius_m)
  movel([0.195893, -1.433129, -2.526477, -0.752783, 1.570796, 1.766690],accel_mss,speed_ms,0,blend_radius_m)
  movel([0.196115, -1.433256, -2.526377, -0.752756, 1.570796, 1.766911],accel_mss,speed_ms,0,blend_radius_m)
  movel([0.196496, -1.433243, -2.526387, -0.752758, 1.570796, 1.767292],accel_mss,speed_ms,0,blend_radius_m)
  movel([0.197345, -1.432020, -2.527347, -0.753023, 1.570796, 1.768141],accel_mss,speed_ms,0,blend_radius_m)
  movel([0.198120, -1.430747, -2.528342, -0.753300, 1.570796, 1.768917],accel_mss,speed_ms,0,blend_radius_m)
  movel([0.197550, -1.435647, -2.524496, -0.752246, 1.570796, 1.768346],accel_mss,speed_ms,0,blend_radius_m)
  movel([0.197168, -1.440466, -2.520679, -0.751244, 1.570796, 1.767964],accel_mss,speed_ms,0,blend_radius_m)
  movel([0.196972, -1.445198, -2.516896, -0.750295, 1.570796, 1.767769],accel_mss,speed_ms,0,blend_radius_m)
  movel([0.196961, -1.449845, -2.513148, -0.749396, 1.570796, 1.767757],accel_mss,speed_ms,0,blend_radius_m)
  movel([0.197034, -1.451836, -2.511531, -0.749021, 1.570796, 1.767830],accel_mss,speed_ms,0,blend_radius_m)
  movel([0.197297, -1.453847, -2.509894, -0.748648, 1.570796, 1.768094],accel_mss,speed_ms,0,blend_radius_m)
  movel([0.197548, -1.454796, -2.509119, -0.748475, 1.570796, 1.768344],accel_mss,speed_ms,0,blend_radius_m)
  movel([0.197903, -1.455671, -2.508402, -0.748316, 1.570796, 1.768699],accel_mss,speed_ms,0,blend_radius_m)
  movel([0.198382, -1.456447, -2.507766, -0.748176, 1.570796, 1.769179],accel_mss,speed_ms,0,blend_radius_m)
  movel([0.199006, -1.457096, -2.507234, -0.748059, 1.570796, 1.769802],accel_mss,speed_ms,0,blend_radius_m)
  movel([0.199534, -1.457451, -2.506942, -0.747996, 1.570796, 1.770330],accel_mss,speed_ms,0,blend_radius_m)
  movel([0.200775, -1.457863, -2.506603, -0.747923, 1.570796, 1.771571],accel_mss,speed_ms,0,blend_radius_m)
  movel([0.201472, -1.457932, -2.506547, -0.747910, 1.570796, 1.772269],accel_mss,speed_ms,0,blend_radius_m)
  movel([0.202982, -1.457834, -2.506627, -0.747928, 1.570796, 1.773778],accel_mss,speed_ms,0,blend_radius_m)
  movel([0.204596, -1.457460, -2.506935, -0.747994, 1.570796, 1.775393],accel_mss,speed_ms,0,blend_radius_m)
  movel([0.206253, -1.456864, -2.507424, -0.748101, 1.570796, 1.777049],accel_mss,speed_ms,0,blend_radius_m)
  movel([0.207892, -1.456095, -2.508055, -0.748239, 1.570796, 1.778689],accel_mss,speed_ms,0,blend_radius_m)
  movel([0.209452, -1.455206, -2.508783, -0.748400, 1.570796, 1.780249],accel_mss,speed_ms,0,blend_radius_m)
  movel([0.210868, -1.454248, -2.509566, -0.748575, 1.570796, 1.781664],accel_mss,speed_ms,0,blend_radius_m)
  speed_ms = 0.005
  movel([0.210868, -1.446215, -2.505864, -0.760310, 1.570796, 1.781664],accel_mss,speed_ms,0,blend_radius_m)
  speed_ms = 0.040
  movel([0.203482, -1.447858, -2.504537, -0.759994, 1.570796, 1.774278],accel_mss,speed_ms,0,blend_radius_m)
  speed_ms = 0.005
  movel([0.203482, -1.455878, -2.508232, -0.748278, 1.570796, 1.774278],accel_mss,speed_ms,0,blend_radius_m)
  speed_ms = 0.025
  movel([0.204628, -1.455055, -2.508907, -0.748427, 1.570796, 1.775424],accel_mss,speed_ms,0,blend_radius_m)
  movel([0.206883, -1.453133, -2.510476, -0.748780, 1.570796, 1.777679],accel_mss,speed_ms,0,blend_radius_m)
  movel([0.207970, -1.452058, -2.511352, -0.748980, 1.570796, 1.778766],accel_mss,speed_ms,0,blend_radius_m)
  movel([0.210012, -1.449734, -2.513237, -0.749417, 1.570796, 1.780809],accel_mss,speed_ms,0,blend_radius_m)
  movel([0.211816, -1.447254, -2.515242, -0.749893, 1.570796, 1.782613],accel_mss,speed_ms,0,blend_radius_m)
  movel([0.212602, -1.445985, -2.516264, -0.750141, 1.570796, 1.783398],accel_mss,speed_ms,0,blend_radius_m)
  movel([0.213295, -1.444708, -2.517289, -0.750392, 1.570796, 1.784092],accel_mss,speed_ms,0,blend_radius_m)
  movel([0.214363, -1.442190, -2.519304, -0.750894, 1.570796, 1.785160],accel_mss,speed_ms,0,blend_radius_m)
  movel([0.214719, -1.440969, -2.520278, -0.751142, 1.570796, 1.785515],accel_mss,speed_ms,0,blend_radius_m)
  movel([0.214938, -1.439793, -2.521214, -0.751382, 1.570796, 1.785734],accel_mss,speed_ms,0,blend_radius_m)
  movel([0.215012, -1.438670, -2.522105, -0.751613, 1.570796, 1.785808],accel_mss,speed_ms,0,blend_radius_m)
  movel([0.214929, -1.437613, -2.522943, -0.751833, 1.570796, 1.785725],accel_mss,speed_ms,0,blend_radius_m)
  movel([0.214652, -1.436380, -2.523918, -0.752091, 1.570796, 1.785448],accel_mss,speed_ms,0,blend_radius_m)
  movel([0.214222, -1.435234, -2.524822, -0.752333, 1.570796, 1.785019],accel_mss,speed_ms,0,blend_radius_m)
  movel([0.213625, -1.434212, -2.525626, -0.752551, 1.570796, 1.784421],accel_mss,speed_ms,0,blend_radius_m)
  movel([0.212845, -1.433355, -2.526300, -0.752734, 1.570796, 1.783641],accel_mss,speed_ms,0,blend_radius_m)
  movel([0.211866, -1.432699, -2.526814, -0.752876, 1.570796, 1.782663],accel_mss,speed_ms,0,blend_radius_m)
  movel([0.210679, -1.432286, -2.527138, -0.752965, 1.570796, 1.781475],accel_mss,speed_ms,0,blend_radius_m)
  movel([0.209266, -1.432153, -2.527242, -0.752994, 1.570796, 1.780062],accel_mss,speed_ms,0,blend_radius_m)
  movel([0.207617, -1.432337, -2.527098, -0.752954, 1.570796, 1.778413],accel_mss,speed_ms,0,blend_radius_m)
  movel([0.206442, -1.432666, -2.526841, -0.752883, 1.570796, 1.777238],accel_mss,speed_ms,0,blend_radius_m)
  movel([0.205265, -1.433168, -2.526447, -0.752774, 1.570796, 1.776061],accel_mss,speed_ms,0,blend_radius_m)
  movel([0.204127, -1.433818, -2.525936, -0.752635, 1.570796, 1.774924],accel_mss,speed_ms,0,blend_radius_m)
  movel([0.203064, -1.434592, -2.525327, -0.752470, 1.570796, 1.773860],accel_mss,speed_ms,0,blend_radius_m)
  movel([0.202112, -1.435466, -2.524639, -0.752284, 1.570796, 1.772908],accel_mss,speed_ms,0,blend_radius_m)
  movel([0.201306, -1.436414, -2.523891, -0.752084, 1.570796, 1.772103],accel_mss,speed_ms,0,blend_radius_m)
  movel([0.200687, -1.437413, -2.523101, -0.751875, 1.570796, 1.771483],accel_mss,speed_ms,0,blend_radius_m)
  movel([0.200284, -1.438440, -2.522288, -0.751661, 1.570796, 1.771080],accel_mss,speed_ms,0,blend_radius_m)
  speed_ms = 0.005
  movel([0.200284, -1.430289, -2.518521, -0.763579, 1.570796, 1.771080],accel_mss,speed_ms,0,blend_radius_m)
  speed_ms = 0.040
  # Splitting Linear movement in 2 (instruction 399: MoveL 378)
  movel([0.226022, -1.445828, -2.506176, -0.760385, 1.570796, 1.796818],accel_mss,speed_ms,0,blend_radius_m)
  movel([0.250548, -1.461966, -2.492971, -0.757452, 1.570796, 1.821345],accel_mss,speed_ms,0,blend_radius_m)
  speed_ms = 0.005
  movel([0.250548, -1.469881, -2.496610, -0.745898, 1.570796, 1.821345],accel_mss,speed_ms,0,blend_radius_m)
  speed_ms = 0.025
  movel([0.248915, -1.475127, -2.492177, -0.745085, 1.570796, 1.819712],accel_mss,speed_ms,0,blend_radius_m)
  movel([0.247903, -1.477733, -2.489960, -0.744696, 1.570796, 1.818699],accel_mss,speed_ms,0,blend_radius_m)
  movel([0.247275, -1.479042, -2.488842, -0.744505, 1.570796, 1.818071],accel_mss,speed_ms,0,blend_radius_m)
  movel([0.246538, -1.480358, -2.487715, -0.744316, 1.570796, 1.817334],accel_mss,speed_ms,0,blend_radius_m)
  movel([0.245619, -1.481729, -2.486539, -0.744121, 1.570796, 1.816415],accel_mss,speed_ms,0,blend_radius_m)
  movel([0.245075, -1.482376, -2.485982, -0.744030, 1.570796, 1.815871],accel_mss,speed_ms,0,blend_radius_m)
  movel([0.244450, -1.482974, -2.485468, -0.743947, 1.570796, 1.815246],accel_mss,speed_ms,0,blend_radius_m)
  movel([0.244631, -1.481745, -2.486525, -0.744119, 1.570796, 1.815427],accel_mss,speed_ms,0,blend_radius_m)
  movel([0.244589, -1.480576, -2.487529, -0.744284, 1.570796, 1.815386],accel_mss,speed_ms,0,blend_radius_m)
  movel([0.244442, -1.480236, -2.487820, -0.744333, 1.570796, 1.815238],accel_mss,speed_ms,0,blend_radius_m)
  movel([0.244241, -1.480186, -2.487863, -0.744340, 1.570796, 1.815038],accel_mss,speed_ms,0,blend_radius_m)
  movel([0.243995, -1.480232, -2.487823, -0.744334, 1.570796, 1.814792],accel_mss,speed_ms,0,blend_radius_m)
  movel([0.243476, -1.480508, -2.487587, -0.744294, 1.570796, 1.814272],accel_mss,speed_ms,0,blend_radius_m)
  movel([0.242718, -1.481121, -2.487061, -0.744207, 1.570796, 1.813514],accel_mss,speed_ms,0,blend_radius_m)
  movel([0.242091, -1.481787, -2.486489, -0.744113, 1.570796, 1.812888],accel_mss,speed_ms,0,blend_radius_m)
  movel([0.241574, -1.482492, -2.485883, -0.744014, 1.570796, 1.812370],accel_mss,speed_ms,0,blend_radius_m)
  movel([0.241140, -1.483224, -2.485252, -0.743912, 1.570796, 1.811937],accel_mss,speed_ms,0,blend_radius_m)
  movel([0.239742, -1.486237, -2.482650, -0.743502, 1.570796, 1.810538],accel_mss,speed_ms,0,blend_radius_m)
  movel([0.238821, -1.487989, -2.481129, -0.743270, 1.570796, 1.809617],accel_mss,speed_ms,0,blend_radius_m)
  movel([0.237775, -1.489717, -2.479626, -0.743046, 1.570796, 1.808571],accel_mss,speed_ms,0,blend_radius_m)
  movel([0.236573, -1.491400, -2.478157, -0.742832, 1.570796, 1.807369],accel_mss,speed_ms,0,blend_radius_m)
  movel([0.235187, -1.493008, -2.476749, -0.742632, 1.570796, 1.805983],accel_mss,speed_ms,0,blend_radius_m)
  movel([0.235719, -1.491621, -2.477963, -0.742804, 1.570796, 1.806515],accel_mss,speed_ms,0,blend_radius_m)
  movel([0.235893, -1.490275, -2.479140, -0.742975, 1.570796, 1.806689],accel_mss,speed_ms,0,blend_radius_m)
  movel([0.235855, -1.489956, -2.479418, -0.743015, 1.570796, 1.806651],accel_mss,speed_ms,0,blend_radius_m)
  movel([0.235680, -1.489723, -2.479621, -0.743045, 1.570796, 1.806476],accel_mss,speed_ms,0,blend_radius_m)
  movel([0.235415, -1.489672, -2.479665, -0.743052, 1.570796, 1.806211],accel_mss,speed_ms,0,blend_radius_m)
  movel([0.235097, -1.489745, -2.479602, -0.743042, 1.570796, 1.805893],accel_mss,speed_ms,0,blend_radius_m)
  movel([0.234445, -1.490107, -2.479286, -0.742996, 1.570796, 1.805241],accel_mss,speed_ms,0,blend_radius_m)
  movel([0.233718, -1.490707, -2.478763, -0.742920, 1.570796, 1.804515],accel_mss,speed_ms,0,blend_radius_m)
  movel([0.233075, -1.491374, -2.478180, -0.742835, 1.570796, 1.803872],accel_mss,speed_ms,0,blend_radius_m)
  movel([0.231981, -1.492833, -2.476902, -0.742654, 1.570796, 1.802777],accel_mss,speed_ms,0,blend_radius_m)
  movel([0.230095, -1.495825, -2.474273, -0.742291, 1.570796, 1.800891],accel_mss,speed_ms,0,blend_radius_m)
  movel([0.228904, -1.497448, -2.472841, -0.742100, 1.570796, 1.799701],accel_mss,speed_ms,0,blend_radius_m)
  movel([0.227597, -1.499022, -2.471448, -0.741919, 1.570796, 1.798393],accel_mss,speed_ms,0,blend_radius_m)
  movel([0.226150, -1.500509, -2.470128, -0.741752, 1.570796, 1.796946],accel_mss,speed_ms,0,blend_radius_m)
  movel([0.224542, -1.501877, -2.468911, -0.741601, 1.570796, 1.795338],accel_mss,speed_ms,0,blend_radius_m)
  movel([0.224933, -1.501130, -2.469576, -0.741683, 1.570796, 1.795730],accel_mss,speed_ms,0,blend_radius_m)
  movel([0.225419, -1.499636, -2.470903, -0.741850, 1.570796, 1.796216],accel_mss,speed_ms,0,blend_radius_m)
  movel([0.225506, -1.498910, -2.471547, -0.741932, 1.570796, 1.796302],accel_mss,speed_ms,0,blend_radius_m)
  movel([0.225462, -1.498597, -2.471825, -0.741968, 1.570796, 1.796258],accel_mss,speed_ms,0,blend_radius_m)
  movel([0.225226, -1.498448, -2.471956, -0.741985, 1.570796, 1.796022],accel_mss,speed_ms,0,blend_radius_m)
  movel([0.224831, -1.498602, -2.471820, -0.741967, 1.570796, 1.795627],accel_mss,speed_ms,0,blend_radius_m)
  movel([0.223904, -1.499218, -2.471274, -0.741897, 1.570796, 1.794700],accel_mss,speed_ms,0,blend_radius_m)
  movel([0.223081, -1.499891, -2.470677, -0.741821, 1.570796, 1.793877],accel_mss,speed_ms,0,blend_radius_m)
  movel([0.221620, -1.501348, -2.469382, -0.741659, 1.570796, 1.792417],accel_mss,speed_ms,0,blend_radius_m)
  movel([0.220203, -1.502845, -2.468048, -0.741496, 1.570796, 1.790999],accel_mss,speed_ms,0,blend_radius_m)
  movel([0.219432, -1.503571, -2.467400, -0.741418, 1.570796, 1.790228],accel_mss,speed_ms,0,blend_radius_m)
  movel([0.218577, -1.504262, -2.466783, -0.741345, 1.570796, 1.789374],accel_mss,speed_ms,0,blend_radius_m)
  movel([0.216386, -1.505790, -2.465414, -0.741185, 1.570796, 1.787182],accel_mss,speed_ms,0,blend_radius_m)
  movel([0.214134, -1.507218, -2.464131, -0.741039, 1.570796, 1.784931],accel_mss,speed_ms,0,blend_radius_m)
  movel([0.211842, -1.508555, -2.462928, -0.740906, 1.570796, 1.782638],accel_mss,speed_ms,0,blend_radius_m)
  movel([0.209522, -1.509818, -2.461789, -0.740782, 1.570796, 1.780318],accel_mss,speed_ms,0,blend_radius_m)
  speed_ms = 0.005
  movel([0.209522, -1.502209, -2.458308, -0.751872, 1.570796, 1.780318],accel_mss,speed_ms,0,blend_radius_m)
  speed_ms = 0.040
  movel([0.196819, -1.480096, -2.477663, -0.754630, 1.570796, 1.767615],accel_mss,speed_ms,0,blend_radius_m)
  speed_ms = 0.005
  movel([0.196819, -1.487875, -2.481229, -0.743285, 1.570796, 1.767615],accel_mss,speed_ms,0,blend_radius_m)
  speed_ms = 0.025
  movel([0.197562, -1.487354, -2.481682, -0.743354, 1.570796, 1.768359],accel_mss,speed_ms,0,blend_radius_m)
  movel([0.198251, -1.486740, -2.482214, -0.743435, 1.570796, 1.769047],accel_mss,speed_ms,0,blend_radius_m)
  movel([0.199538, -1.485344, -2.483423, -0.743622, 1.570796, 1.770334],accel_mss,speed_ms,0,blend_radius_m)
  movel([0.200816, -1.483905, -2.484666, -0.743818, 1.570796, 1.771613],accel_mss,speed_ms,0,blend_radius_m)
  movel([0.201499, -1.483237, -2.485242, -0.743911, 1.570796, 1.772295],accel_mss,speed_ms,0,blend_radius_m)
  movel([0.202232, -1.482640, -2.485755, -0.743993, 1.570796, 1.773028],accel_mss,speed_ms,0,blend_radius_m)
  movel([0.202799, -1.482277, -2.486068, -0.744044, 1.570796, 1.773595],accel_mss,speed_ms,0,blend_radius_m)
  movel([0.203252, -1.482081, -2.486236, -0.744072, 1.570796, 1.774048],accel_mss,speed_ms,0,blend_radius_m)
  movel([0.203602, -1.482031, -2.486279, -0.744079, 1.570796, 1.774398],accel_mss,speed_ms,0,blend_radius_m)
  movel([0.203862, -1.482110, -2.486211, -0.744068, 1.570796, 1.774658],accel_mss,speed_ms,0,blend_radius_m)
  movel([0.204140, -1.482590, -2.485799, -0.744000, 1.570796, 1.774937],accel_mss,speed_ms,0,blend_radius_m)
  movel([0.204170, -1.483374, -2.485124, -0.743892, 1.570796, 1.774967],accel_mss,speed_ms,0,blend_radius_m)
  movel([0.203796, -1.485290, -2.483469, -0.743630, 1.570796, 1.774592],accel_mss,speed_ms,0,blend_radius_m)
  movel([0.203381, -1.486729, -2.482224, -0.743437, 1.570796, 1.774178],accel_mss,speed_ms,0,blend_radius_m)
  movel([0.204765, -1.485340, -2.483426, -0.743623, 1.570796, 1.775561],accel_mss,speed_ms,0,blend_radius_m)
  movel([0.205870, -1.483929, -2.484645, -0.743815, 1.570796, 1.776666],accel_mss,speed_ms,0,blend_radius_m)
  movel([0.206769, -1.482495, -2.485881, -0.744014, 1.570796, 1.777566],accel_mss,speed_ms,0,blend_radius_m)
  movel([0.207529, -1.481043, -2.487128, -0.744218, 1.570796, 1.778325],accel_mss,speed_ms,0,blend_radius_m)
  movel([0.209674, -1.476600, -2.490925, -0.744864, 1.570796, 1.780470],accel_mss,speed_ms,0,blend_radius_m)
  movel([0.210576, -1.475098, -2.492202, -0.745089, 1.570796, 1.781373],accel_mss,speed_ms,0,blend_radius_m)
  movel([0.211039, -1.474525, -2.492689, -0.745176, 1.570796, 1.781835],accel_mss,speed_ms,0,blend_radius_m)
  movel([0.211471, -1.474208, -2.492957, -0.745224, 1.570796, 1.782267],accel_mss,speed_ms,0,blend_radius_m)
  movel([0.211866, -1.474107, -2.493043, -0.745240, 1.570796, 1.782662],accel_mss,speed_ms,0,blend_radius_m)
  movel([0.212214, -1.474183, -2.492978, -0.745228, 1.570796, 1.783010],accel_mss,speed_ms,0,blend_radius_m)
  movel([0.212510, -1.474394, -2.492800, -0.745196, 1.570796, 1.783307],accel_mss,speed_ms,0,blend_radius_m)
  movel([0.212743, -1.474700, -2.492540, -0.745149, 1.570796, 1.783540],accel_mss,speed_ms,0,blend_radius_m)
  movel([0.212996, -1.475436, -2.491915, -0.745038, 1.570796, 1.783792],accel_mss,speed_ms,0,blend_radius_m)
  movel([0.212944, -1.476262, -2.491213, -0.744914, 1.570796, 1.783741],accel_mss,speed_ms,0,blend_radius_m)
  movel([0.212689, -1.477339, -2.490296, -0.744754, 1.570796, 1.783486],accel_mss,speed_ms,0,blend_radius_m)
  movel([0.212081, -1.479330, -2.488596, -0.744463, 1.570796, 1.782877],accel_mss,speed_ms,0,blend_radius_m)
  movel([0.213725, -1.476345, -2.491142, -0.744902, 1.570796, 1.784521],accel_mss,speed_ms,0,blend_radius_m)
  movel([0.214406, -1.474837, -2.492424, -0.745128, 1.570796, 1.785202],accel_mss,speed_ms,0,blend_radius_m)
  movel([0.215476, -1.471810, -2.494985, -0.745594, 1.570796, 1.786273],accel_mss,speed_ms,0,blend_radius_m)
  movel([0.215858, -1.470306, -2.496252, -0.745831, 1.570796, 1.786655],accel_mss,speed_ms,0,blend_radius_m)
  movel([0.216308, -1.467345, -2.498737, -0.746307, 1.570796, 1.787104],accel_mss,speed_ms,0,blend_radius_m)
  speed_ms = 0.005
  movel([0.216308, -1.459410, -2.495089, -0.757890, 1.570796, 1.787104],accel_mss,speed_ms,0,blend_radius_m)
  speed_ms = 0.040
  movel([0.203967, -1.469939, -2.486301, -0.756149, 1.570796, 1.774764],accel_mss,speed_ms,0,blend_radius_m)
  speed_ms = 0.005
  movel([0.203967, -1.477794, -2.489907, -0.744687, 1.570796, 1.774764],accel_mss,speed_ms,0,blend_radius_m)
  speed_ms = 0.025
  movel([0.202357, -1.479358, -2.488572, -0.744459, 1.570796, 1.773154],accel_mss,speed_ms,0,blend_radius_m)
  movel([0.200852, -1.480985, -2.487178, -0.744226, 1.570796, 1.771649],accel_mss,speed_ms,0,blend_radius_m)
  movel([0.197910, -1.484267, -2.484354, -0.743769, 1.570796, 1.768706],accel_mss,speed_ms,0,blend_radius_m)
  movel([0.196330, -1.485850, -2.482985, -0.743554, 1.570796, 1.767126],accel_mss,speed_ms,0,blend_radius_m)
  movel([0.194623, -1.487323, -2.481708, -0.743358, 1.570796, 1.765420],accel_mss,speed_ms,0,blend_radius_m)
  movel([0.192788, -1.488597, -2.480601, -0.743191, 1.570796, 1.763584],accel_mss,speed_ms,0,blend_radius_m)
  movel([0.191824, -1.489134, -2.480134, -0.743121, 1.570796, 1.762620],accel_mss,speed_ms,0,blend_radius_m)
  movel([0.190828, -1.489589, -2.479737, -0.743062, 1.570796, 1.761625],accel_mss,speed_ms,0,blend_radius_m)
  movel([0.191579, -1.489124, -2.480143, -0.743122, 1.570796, 1.762375],accel_mss,speed_ms,0,blend_radius_m)
  movel([0.192409, -1.488355, -2.480812, -0.743222, 1.570796, 1.763206],accel_mss,speed_ms,0,blend_radius_m)
  movel([0.193220, -1.487397, -2.481644, -0.743348, 1.570796, 1.764017],accel_mss,speed_ms,0,blend_radius_m)
  movel([0.193900, -1.486371, -2.482534, -0.743484, 1.570796, 1.764697],accel_mss,speed_ms,0,blend_radius_m)
  movel([0.194346, -1.485390, -2.483383, -0.743616, 1.570796, 1.765142],accel_mss,speed_ms,0,blend_radius_m)
  movel([0.194445, -1.484957, -2.483758, -0.743675, 1.570796, 1.765241],accel_mss,speed_ms,0,blend_radius_m)
  movel([0.194446, -1.484579, -2.484084, -0.743726, 1.570796, 1.765242],accel_mss,speed_ms,0,blend_radius_m)
  movel([0.194335, -1.484271, -2.484349, -0.743768, 1.570796, 1.765131],accel_mss,speed_ms,0,blend_radius_m)
  movel([0.194095, -1.484052, -2.484539, -0.743798, 1.570796, 1.764892],accel_mss,speed_ms,0,blend_radius_m)
  movel([0.193719, -1.483933, -2.484642, -0.743815, 1.570796, 1.764515],accel_mss,speed_ms,0,blend_radius_m)
  movel([0.193186, -1.483930, -2.484644, -0.743815, 1.570796, 1.763983],accel_mss,speed_ms,0,blend_radius_m)
  movel([0.192285, -1.484188, -2.484422, -0.743780, 1.570796, 1.763081],accel_mss,speed_ms,0,blend_radius_m)
  movel([0.188439, -1.486014, -2.482843, -0.743532, 1.570796, 1.759235],accel_mss,speed_ms,0,blend_radius_m)
  movel([0.186816, -1.486644, -2.482297, -0.743448, 1.570796, 1.757612],accel_mss,speed_ms,0,blend_radius_m)
  movel([0.185169, -1.487165, -2.481845, -0.743379, 1.570796, 1.755966],accel_mss,speed_ms,0,blend_radius_m)
  movel([0.183557, -1.487534, -2.481525, -0.743330, 1.570796, 1.754353],accel_mss,speed_ms,0,blend_radius_m)
  movel([0.182035, -1.487700, -2.481381, -0.743308, 1.570796, 1.752832],accel_mss,speed_ms,0,blend_radius_m)
  movel([0.180660, -1.487617, -2.481453, -0.743319, 1.570796, 1.751456],accel_mss,speed_ms,0,blend_radius_m)
  movel([0.179490, -1.487233, -2.481787, -0.743370, 1.570796, 1.750286],accel_mss,speed_ms,0,blend_radius_m)
  movel([0.179876, -1.487293, -2.481734, -0.743362, 1.570796, 1.750672],accel_mss,speed_ms,0,blend_radius_m)
  movel([0.180416, -1.487196, -2.481819, -0.743375, 1.570796, 1.751212],accel_mss,speed_ms,0,blend_radius_m)
  movel([0.181762, -1.486673, -2.482272, -0.743444, 1.570796, 1.752559],accel_mss,speed_ms,0,blend_radius_m)
  movel([0.183120, -1.485954, -2.482895, -0.743540, 1.570796, 1.753916],accel_mss,speed_ms,0,blend_radius_m)
  movel([0.184076, -1.485335, -2.483431, -0.743623, 1.570796, 1.754872],accel_mss,speed_ms,0,blend_radius_m)
  movel([0.184667, -1.484805, -2.483888, -0.743695, 1.570796, 1.755463],accel_mss,speed_ms,0,blend_radius_m)
  movel([0.184924, -1.484401, -2.484237, -0.743750, 1.570796, 1.755721],accel_mss,speed_ms,0,blend_radius_m)
  movel([0.184902, -1.484103, -2.484495, -0.743791, 1.570796, 1.755698],accel_mss,speed_ms,0,blend_radius_m)
  movel([0.184660, -1.483894, -2.484675, -0.743820, 1.570796, 1.755456],accel_mss,speed_ms,0,blend_radius_m)
  movel([0.183750, -1.483671, -2.484867, -0.743851, 1.570796, 1.754547],accel_mss,speed_ms,0,blend_radius_m)
  movel([0.182663, -1.483593, -2.484935, -0.743861, 1.570796, 1.753459],accel_mss,speed_ms,0,blend_radius_m)
  movel([0.180191, -1.483411, -2.485092, -0.743886, 1.570796, 1.750987],accel_mss,speed_ms,0,blend_radius_m)
  movel([0.177769, -1.483014, -2.485433, -0.743941, 1.570796, 1.748566],accel_mss,speed_ms,0,blend_radius_m)
  movel([0.176653, -1.482683, -2.485718, -0.743987, 1.570796, 1.747450],accel_mss,speed_ms,0,blend_radius_m)
  movel([0.175642, -1.482234, -2.486105, -0.744050, 1.570796, 1.746438],accel_mss,speed_ms,0,blend_radius_m)
  movel([0.174767, -1.481645, -2.486611, -0.744133, 1.570796, 1.745564],accel_mss,speed_ms,0,blend_radius_m)
  movel([0.174060, -1.480894, -2.487256, -0.744239, 1.570796, 1.744856],accel_mss,speed_ms,0,blend_radius_m)
  movel([0.175538, -1.480993, -2.487171, -0.744225, 1.570796, 1.746334],accel_mss,speed_ms,0,blend_radius_m)
  movel([0.176381, -1.480869, -2.487277, -0.744243, 1.570796, 1.747178],accel_mss,speed_ms,0,blend_radius_m)
  movel([0.176773, -1.480722, -2.487404, -0.744264, 1.570796, 1.747569],accel_mss,speed_ms,0,blend_radius_m)
  movel([0.177126, -1.480497, -2.487596, -0.744296, 1.570796, 1.747922],accel_mss,speed_ms,0,blend_radius_m)
  movel([0.177294, -1.480284, -2.487779, -0.744326, 1.570796, 1.748090],accel_mss,speed_ms,0,blend_radius_m)
  movel([0.177323, -1.480039, -2.487989, -0.744361, 1.570796, 1.748119],accel_mss,speed_ms,0,blend_radius_m)
  movel([0.177039, -1.479479, -2.488468, -0.744442, 1.570796, 1.747835],accel_mss,speed_ms,0,blend_radius_m)
  movel([0.176400, -1.478861, -2.488996, -0.744531, 1.570796, 1.747196],accel_mss,speed_ms,0,blend_radius_m)
  movel([0.175537, -1.478226, -2.489539, -0.744624, 1.570796, 1.746333],accel_mss,speed_ms,0,blend_radius_m)
  movel([0.172444, -1.476369, -2.491122, -0.744898, 1.570796, 1.743240],accel_mss,speed_ms,0,blend_radius_m)
  movel([0.171365, -1.475489, -2.491870, -0.745030, 1.570796, 1.742161],accel_mss,speed_ms,0,blend_radius_m)
  movel([0.170434, -1.474480, -2.492726, -0.745183, 1.570796, 1.741230],accel_mss,speed_ms,0,blend_radius_m)
  movel([0.169729, -1.473321, -2.493708, -0.745360, 1.570796, 1.740525],accel_mss,speed_ms,0,blend_radius_m)
  movel([0.169319, -1.471989, -2.494833, -0.745566, 1.570796, 1.740116],accel_mss,speed_ms,0,blend_radius_m)
  movel([0.170298, -1.472876, -2.494084, -0.745428, 1.570796, 1.741095],accel_mss,speed_ms,0,blend_radius_m)
  movel([0.170948, -1.473235, -2.493780, -0.745373, 1.570796, 1.741744],accel_mss,speed_ms,0,blend_radius_m)
  movel([0.171629, -1.473334, -2.493697, -0.745358, 1.570796, 1.742426],accel_mss,speed_ms,0,blend_radius_m)
  movel([0.172340, -1.473125, -2.493874, -0.745390, 1.570796, 1.743136],accel_mss,speed_ms,0,blend_radius_m)
  movel([0.172820, -1.472727, -2.494210, -0.745452, 1.570796, 1.743617],accel_mss,speed_ms,0,blend_radius_m)
  movel([0.173042, -1.472211, -2.494647, -0.745532, 1.570796, 1.743838],accel_mss,speed_ms,0,blend_radius_m)
  movel([0.172979, -1.471642, -2.495127, -0.745620, 1.570796, 1.743775],accel_mss,speed_ms,0,blend_radius_m)
  movel([0.172084, -1.468800, -2.497518, -0.746071, 1.570796, 1.742880],accel_mss,speed_ms,0,blend_radius_m)
  movel([0.171564, -1.465851, -2.499985, -0.746552, 1.570796, 1.742360],accel_mss,speed_ms,0,blend_radius_m)
  movel([0.171476, -1.464307, -2.501272, -0.746809, 1.570796, 1.742272],accel_mss,speed_ms,0,blend_radius_m)
  movel([0.171518, -1.462701, -2.502607, -0.747081, 1.570796, 1.742314],accel_mss,speed_ms,0,blend_radius_m)
  movel([0.171704, -1.461019, -2.504000, -0.747369, 1.570796, 1.742500],accel_mss,speed_ms,0,blend_radius_m)
  movel([0.172044, -1.459251, -2.505461, -0.747677, 1.570796, 1.742841],accel_mss,speed_ms,0,blend_radius_m)
  speed_ms = 0.005
  movel([0.172044, -1.451255, -2.501779, -0.759355, 1.570796, 1.742841],accel_mss,speed_ms,0,blend_radius_m)
  speed_ms = 0.040
  movel([0.151825, -1.436811, -2.513384, -0.762194, 1.570796, 1.722621],accel_mss,speed_ms,0,blend_radius_m)
  speed_ms = 0.005
  movel([0.151825, -1.444914, -2.517124, -0.750351, 1.570796, 1.722621],accel_mss,speed_ms,0,blend_radius_m)
  speed_ms = 0.025
  movel([0.154240, -1.442524, -2.519038, -0.750827, 1.570796, 1.725037],accel_mss,speed_ms,0,blend_radius_m)
  movel([0.156589, -1.440083, -2.520984, -0.751323, 1.570796, 1.727385],accel_mss,speed_ms,0,blend_radius_m)
  movel([0.161126, -1.435047, -2.524969, -0.752373, 1.570796, 1.731922],accel_mss,speed_ms,0,blend_radius_m)
  movel([0.165440, -1.429821, -2.529065, -0.753503, 1.570796, 1.736237],accel_mss,speed_ms,0,blend_radius_m)
  movel([0.169523, -1.424423, -2.533252, -0.754713, 1.570796, 1.740319],accel_mss,speed_ms,0,blend_radius_m)
  movel([0.173366, -1.418868, -2.537516, -0.756005, 1.570796, 1.744162],accel_mss,speed_ms,0,blend_radius_m)
  movel([0.176958, -1.413175, -2.541839, -0.757375, 1.570796, 1.747754],accel_mss,speed_ms,0,blend_radius_m)
  movel([0.180289, -1.407364, -2.546201, -0.758824, 1.570796, 1.751085],accel_mss,speed_ms,0,blend_radius_m)
  movel([0.183348, -1.401453, -2.550588, -0.760348, 1.570796, 1.754145],accel_mss,speed_ms,0,blend_radius_m)
  movel([0.186122, -1.395467, -2.554978, -0.761944, 1.570796, 1.756918],accel_mss,speed_ms,0,blend_radius_m)
  movel([0.188597, -1.389426, -2.559356, -0.763607, 1.570796, 1.759393],accel_mss,speed_ms,0,blend_radius_m)
  movel([0.190758, -1.383354, -2.563703, -0.765332, 1.570796, 1.761555],accel_mss,speed_ms,0,blend_radius_m)
  movel([0.192589, -1.377277, -2.568001, -0.767111, 1.570796, 1.763386],accel_mss,speed_ms,0,blend_radius_m)
  movel([0.194081, -1.371218, -2.572234, -0.768937, 1.570796, 1.764877],accel_mss,speed_ms,0,blend_radius_m)
  movel([0.195210, -1.365208, -2.576382, -0.770800, 1.570796, 1.766006],accel_mss,speed_ms,0,blend_radius_m)
  movel([0.195963, -1.359275, -2.580426, -0.772689, 1.570796, 1.766760],accel_mss,speed_ms,0,blend_radius_m)
  movel([0.196494, -1.350524, -2.586301, -0.775564, 1.570796, 1.767290],accel_mss,speed_ms,0,blend_radius_m)
  movel([0.196790, -1.349012, -2.587306, -0.776071, 1.570796, 1.767586],accel_mss,speed_ms,0,blend_radius_m)
  movel([0.197348, -1.347459, -2.588334, -0.776596, 1.570796, 1.768145],accel_mss,speed_ms,0,blend_radius_m)
  movel([0.198479, -1.345323, -2.589743, -0.777323, 1.570796, 1.769276],accel_mss,speed_ms,0,blend_radius_m)
  movel([0.199662, -1.343710, -2.590803, -0.777876, 1.570796, 1.770458],accel_mss,speed_ms,0,blend_radius_m)
  movel([0.200265, -1.343088, -2.591211, -0.778090, 1.570796, 1.771062],accel_mss,speed_ms,0,blend_radius_m)
  movel([0.201493, -1.342180, -2.591805, -0.778404, 1.570796, 1.772289],accel_mss,speed_ms,0,blend_radius_m)
  movel([0.202108, -1.341887, -2.591997, -0.778505, 1.570796, 1.772905],accel_mss,speed_ms,0,blend_radius_m)
  movel([0.203343, -1.341590, -2.592191, -0.778608, 1.570796, 1.774139],accel_mss,speed_ms,0,blend_radius_m)
  movel([0.204563, -1.341640, -2.592158, -0.778591, 1.570796, 1.775359],accel_mss,speed_ms,0,blend_radius_m)
  movel([0.205753, -1.341991, -2.591929, -0.778469, 1.570796, 1.776550],accel_mss,speed_ms,0,blend_radius_m)
  movel([0.206901, -1.342599, -2.591531, -0.778259, 1.570796, 1.777697],accel_mss,speed_ms,0,blend_radius_m)
  movel([0.207989, -1.343412, -2.590998, -0.777978, 1.570796, 1.778786],accel_mss,speed_ms,0,blend_radius_m)
  movel([0.209006, -1.344388, -2.590358, -0.777643, 1.570796, 1.779803],accel_mss,speed_ms,0,blend_radius_m)
  movel([0.210767, -1.346625, -2.588885, -0.776879, 1.570796, 1.781563],accel_mss,speed_ms,0,blend_radius_m)
  movel([0.212076, -1.348935, -2.587357, -0.776097, 1.570796, 1.782872],accel_mss,speed_ms,0,blend_radius_m)
  movel([0.212839, -1.350935, -2.586028, -0.775426, 1.570796, 1.783635],accel_mss,speed_ms,0,blend_radius_m)
  movel([0.213362, -1.353450, -2.584348, -0.774590, 1.570796, 1.784158],accel_mss,speed_ms,0,blend_radius_m)
  movel([0.213674, -1.356064, -2.582594, -0.773731, 1.570796, 1.784470],accel_mss,speed_ms,0,blend_radius_m)
  movel([0.213879, -1.361461, -2.578941, -0.771987, 1.570796, 1.784676],accel_mss,speed_ms,0,blend_radius_m)
  movel([0.213867, -1.366895, -2.575222, -0.770272, 1.570796, 1.784663],accel_mss,speed_ms,0,blend_radius_m)
  movel([0.214034, -1.372144, -2.571590, -0.768654, 1.570796, 1.784831],accel_mss,speed_ms,0,blend_radius_m)
  movel([0.214513, -1.376684, -2.568418, -0.767287, 1.570796, 1.785309],accel_mss,speed_ms,0,blend_radius_m)
  movel([0.214993, -1.378819, -2.566915, -0.766654, 1.570796, 1.785789],accel_mss,speed_ms,0,blend_radius_m)
  movel([0.215765, -1.380782, -2.565529, -0.766078, 1.570796, 1.786562],accel_mss,speed_ms,0,blend_radius_m)
  movel([0.216300, -1.381583, -2.564961, -0.765845, 1.570796, 1.787097],accel_mss,speed_ms,0,blend_radius_m)
  movel([0.216675, -1.381886, -2.564746, -0.765757, 1.570796, 1.787471],accel_mss,speed_ms,0,blend_radius_m)
  movel([0.217149, -1.382076, -2.564612, -0.765701, 1.570796, 1.787945],accel_mss,speed_ms,0,blend_radius_m)
  movel([0.217882, -1.382109, -2.564588, -0.765692, 1.570796, 1.788679],accel_mss,speed_ms,0,blend_radius_m)
  movel([0.218690, -1.381941, -2.564707, -0.765741, 1.570796, 1.789486],accel_mss,speed_ms,0,blend_radius_m)
  movel([0.220372, -1.381231, -2.565211, -0.765947, 1.570796, 1.791168],accel_mss,speed_ms,0,blend_radius_m)
  movel([0.222255, -1.380188, -2.565949, -0.766252, 1.570796, 1.793051],accel_mss,speed_ms,0,blend_radius_m)
  movel([0.224077, -1.379029, -2.566768, -0.766593, 1.570796, 1.794873],accel_mss,speed_ms,0,blend_radius_m)
  movel([0.227586, -1.376448, -2.568583, -0.767357, 1.570796, 1.798382],accel_mss,speed_ms,0,blend_radius_m)
  movel([0.234441, -1.370917, -2.572443, -0.769029, 1.570796, 1.805237],accel_mss,speed_ms,0,blend_radius_m)
  movel([0.237750, -1.368433, -2.574162, -0.769794, 1.570796, 1.808546],accel_mss,speed_ms,0,blend_radius_m)
  movel([0.239656, -1.367159, -2.575041, -0.770189, 1.570796, 1.810452],accel_mss,speed_ms,0,blend_radius_m)
  movel([0.241539, -1.366103, -2.575767, -0.770519, 1.570796, 1.812335],accel_mss,speed_ms,0,blend_radius_m)
  movel([0.242428, -1.365711, -2.576036, -0.770642, 1.570796, 1.813224],accel_mss,speed_ms,0,blend_radius_m)
  movel([0.243258, -1.365440, -2.576222, -0.770727, 1.570796, 1.814055],accel_mss,speed_ms,0,blend_radius_m)
  movel([0.244011, -1.365311, -2.576311, -0.770767, 1.570796, 1.814807],accel_mss,speed_ms,0,blend_radius_m)
  movel([0.244669, -1.365349, -2.576285, -0.770755, 1.570796, 1.815466],accel_mss,speed_ms,0,blend_radius_m)
  movel([0.245214, -1.365572, -2.576132, -0.770685, 1.570796, 1.816010],accel_mss,speed_ms,0,blend_radius_m)
  movel([0.245629, -1.366002, -2.575836, -0.770551, 1.570796, 1.816425],accel_mss,speed_ms,0,blend_radius_m)
  movel([0.245895, -1.366663, -2.575382, -0.770344, 1.570796, 1.816692],accel_mss,speed_ms,0,blend_radius_m)
  movel([0.245995, -1.367575, -2.574754, -0.770060, 1.570796, 1.816791],accel_mss,speed_ms,0,blend_radius_m)
  movel([0.245926, -1.369271, -2.573583, -0.769535, 1.570796, 1.816722],accel_mss,speed_ms,0,blend_radius_m)
  movel([0.245685, -1.370972, -2.572405, -0.769012, 1.570796, 1.816482],accel_mss,speed_ms,0,blend_radius_m)
  movel([0.245286, -1.372672, -2.571223, -0.768494, 1.570796, 1.816082],accel_mss,speed_ms,0,blend_radius_m)
  movel([0.244737, -1.374373, -2.570037, -0.767980, 1.570796, 1.815533],accel_mss,speed_ms,0,blend_radius_m)
  movel([0.244047, -1.376063, -2.568854, -0.767473, 1.570796, 1.814843],accel_mss,speed_ms,0,blend_radius_m)
  movel([0.243226, -1.377742, -2.567675, -0.766973, 1.570796, 1.814022],accel_mss,speed_ms,0,blend_radius_m)
  movel([0.242283, -1.379405, -2.566502, -0.766482, 1.570796, 1.813079],accel_mss,speed_ms,0,blend_radius_m)
  movel([0.241228, -1.381051, -2.565339, -0.766000, 1.570796, 1.812025],accel_mss,speed_ms,0,blend_radius_m)
  movel([0.238823, -1.384267, -2.563053, -0.765069, 1.570796, 1.809619],accel_mss,speed_ms,0,blend_radius_m)
  movel([0.236079, -1.387365, -2.560838, -0.764186, 1.570796, 1.806876],accel_mss,speed_ms,0,blend_radius_m)
  movel([0.233067, -1.390316, -2.558714, -0.763358, 1.570796, 1.803864],accel_mss,speed_ms,0,blend_radius_m)
  movel([0.229862, -1.393094, -2.556704, -0.762591, 1.570796, 1.800658],accel_mss,speed_ms,0,blend_radius_m)
  movel([0.222508, -1.399044, -2.552361, -0.760984, 1.570796, 1.793304],accel_mss,speed_ms,0,blend_radius_m)
  movel([0.218667, -1.401838, -2.550304, -0.760247, 1.570796, 1.789464],accel_mss,speed_ms,0,blend_radius_m)
  movel([0.216733, -1.403088, -2.549380, -0.759921, 1.570796, 1.787529],accel_mss,speed_ms,0,blend_radius_m)
  movel([0.214796, -1.404202, -2.548554, -0.759633, 1.570796, 1.785592],accel_mss,speed_ms,0,blend_radius_m)
  movel([0.213553, -1.404821, -2.548095, -0.759473, 1.570796, 1.784349],accel_mss,speed_ms,0,blend_radius_m)
  movel([0.212326, -1.405328, -2.547718, -0.759343, 1.570796, 1.783122],accel_mss,speed_ms,0,blend_radius_m)
  movel([0.211125, -1.405711, -2.547433, -0.759245, 1.570796, 1.781921],accel_mss,speed_ms,0,blend_radius_m)
  movel([0.209962, -1.405955, -2.547252, -0.759182, 1.570796, 1.780759],accel_mss,speed_ms,0,blend_radius_m)
  movel([0.208851, -1.406047, -2.547183, -0.759159, 1.570796, 1.779648],accel_mss,speed_ms,0,blend_radius_m)
  movel([0.207802, -1.405974, -2.547237, -0.759178, 1.570796, 1.778598],accel_mss,speed_ms,0,blend_radius_m)
  movel([0.206829, -1.405718, -2.547428, -0.759243, 1.570796, 1.777625],accel_mss,speed_ms,0,blend_radius_m)
  movel([0.205941, -1.405265, -2.547765, -0.759359, 1.570796, 1.776738],accel_mss,speed_ms,0,blend_radius_m)
  movel([0.205185, -1.404617, -2.548246, -0.759526, 1.570796, 1.775981],accel_mss,speed_ms,0,blend_radius_m)
  movel([0.204601, -1.403846, -2.548818, -0.759725, 1.570796, 1.775397],accel_mss,speed_ms,0,blend_radius_m)
  movel([0.202831, -1.400317, -2.551425, -0.760647, 1.570796, 1.773628],accel_mss,speed_ms,0,blend_radius_m)
  movel([0.202235, -1.399525, -2.552007, -0.760856, 1.570796, 1.773031],accel_mss,speed_ms,0,blend_radius_m)
  movel([0.201456, -1.398853, -2.552501, -0.761035, 1.570796, 1.772252],accel_mss,speed_ms,0,blend_radius_m)
  movel([0.201068, -1.398710, -2.552607, -0.761073, 1.570796, 1.771865],accel_mss,speed_ms,0,blend_radius_m)
  movel([0.200840, -1.398888, -2.552475, -0.761025, 1.570796, 1.771636],accel_mss,speed_ms,0,blend_radius_m)
  movel([0.200488, -1.399389, -2.552108, -0.760892, 1.570796, 1.771284],accel_mss,speed_ms,0,blend_radius_m)
  movel([0.199472, -1.401190, -2.550782, -0.760417, 1.570796, 1.770269],accel_mss,speed_ms,0,blend_radius_m)
  movel([0.196728, -1.406737, -2.546669, -0.758983, 1.570796, 1.767524],accel_mss,speed_ms,0,blend_radius_m)
  movel([0.192310, -1.416029, -2.539678, -0.756682, 1.570796, 1.763107],accel_mss,speed_ms,0,blend_radius_m)
  movel([0.189482, -1.420817, -2.536026, -0.755546, 1.570796, 1.760279],accel_mss,speed_ms,0,blend_radius_m)
  movel([0.186452, -1.425525, -2.532401, -0.754463, 1.570796, 1.757248],accel_mss,speed_ms,0,blend_radius_m)
  movel([0.183244, -1.430153, -2.528806, -0.753430, 1.570796, 1.754040],accel_mss,speed_ms,0,blend_radius_m)
  movel([0.179892, -1.434694, -2.525247, -0.752448, 1.570796, 1.750689],accel_mss,speed_ms,0,blend_radius_m)
  movel([0.175483, -1.440419, -2.520716, -0.751254, 1.570796, 1.746279],accel_mss,speed_ms,0,blend_radius_m)
  movel([0.170963, -1.446071, -2.516194, -0.750124, 1.570796, 1.741759],accel_mss,speed_ms,0,blend_radius_m)
  movel([0.166313, -1.451614, -2.511712, -0.749063, 1.570796, 1.737109],accel_mss,speed_ms,0,blend_radius_m)
  movel([0.161506, -1.457009, -2.507305, -0.748075, 1.570796, 1.732303],accel_mss,speed_ms,0,blend_radius_m)
  movel([0.156524, -1.462217, -2.503009, -0.747164, 1.570796, 1.727320],accel_mss,speed_ms,0,blend_radius_m)
  movel([0.153962, -1.464740, -2.500912, -0.746737, 1.570796, 1.724758],accel_mss,speed_ms,0,blend_radius_m)
  movel([0.151344, -1.467204, -2.498855, -0.746330, 1.570796, 1.722140],accel_mss,speed_ms,0,blend_radius_m)
  movel([0.148670, -1.469604, -2.496842, -0.745942, 1.570796, 1.719466],accel_mss,speed_ms,0,blend_radius_m)
  movel([0.145939, -1.471935, -2.494880, -0.745575, 1.570796, 1.716735],accel_mss,speed_ms,0,blend_radius_m)
  movel([0.143145, -1.474196, -2.492967, -0.745226, 1.570796, 1.713941],accel_mss,speed_ms,0,blend_radius_m)
  movel([0.140284, -1.476379, -2.491113, -0.744897, 1.570796, 1.711080],accel_mss,speed_ms,0,blend_radius_m)
  movel([0.136811, -1.478871, -2.488988, -0.744530, 1.570796, 1.707607],accel_mss,speed_ms,0,blend_radius_m)
  movel([0.135028, -1.480026, -2.487999, -0.744363, 1.570796, 1.705824],accel_mss,speed_ms,0,blend_radius_m)
  movel([0.131882, -1.481769, -2.486504, -0.744115, 1.570796, 1.702679],accel_mss,speed_ms,0,blend_radius_m)
  movel([0.130288, -1.482499, -2.485877, -0.744013, 1.570796, 1.701084],accel_mss,speed_ms,0,blend_radius_m)
  movel([0.128742, -1.482965, -2.485476, -0.743948, 1.570796, 1.699538],accel_mss,speed_ms,0,blend_radius_m)
  movel([0.128090, -1.483003, -2.485443, -0.743943, 1.570796, 1.698886],accel_mss,speed_ms,0,blend_radius_m)
  movel([0.127568, -1.482862, -2.485564, -0.743963, 1.570796, 1.698364],accel_mss,speed_ms,0,blend_radius_m)
  movel([0.128271, -1.481450, -2.486778, -0.744160, 1.570796, 1.699067],accel_mss,speed_ms,0,blend_radius_m)
  movel([0.128763, -1.480037, -2.487991, -0.744362, 1.570796, 1.699560],accel_mss,speed_ms,0,blend_radius_m)
  movel([0.128867, -1.479378, -2.488554, -0.744456, 1.570796, 1.699663],accel_mss,speed_ms,0,blend_radius_m)
  movel([0.128840, -1.478778, -2.489068, -0.744543, 1.570796, 1.699636],accel_mss,speed_ms,0,blend_radius_m)
  movel([0.128658, -1.478254, -2.489515, -0.744620, 1.570796, 1.699455],accel_mss,speed_ms,0,blend_radius_m)
  movel([0.128291, -1.477830, -2.489877, -0.744682, 1.570796, 1.699087],accel_mss,speed_ms,0,blend_radius_m)
  movel([0.127035, -1.477109, -2.490492, -0.744788, 1.570796, 1.697831],accel_mss,speed_ms,0,blend_radius_m)
  movel([0.126724, -1.476739, -2.490807, -0.744843, 1.570796, 1.697520],accel_mss,speed_ms,0,blend_radius_m)
  movel([0.126553, -1.476289, -2.491190, -0.744910, 1.570796, 1.697350],accel_mss,speed_ms,0,blend_radius_m)
  movel([0.126566, -1.475215, -2.492103, -0.745071, 1.570796, 1.697363],accel_mss,speed_ms,0,blend_radius_m)
  movel([0.126919, -1.474006, -2.493128, -0.745255, 1.570796, 1.697715],accel_mss,speed_ms,0,blend_radius_m)
  movel([0.127458, -1.472786, -2.494160, -0.745442, 1.570796, 1.698254],accel_mss,speed_ms,0,blend_radius_m)
  movel([0.129320, -1.469134, -2.497237, -0.746018, 1.570796, 1.700116],accel_mss,speed_ms,0,blend_radius_m)
  movel([0.131423, -1.465462, -2.500310, -0.746617, 1.570796, 1.702219],accel_mss,speed_ms,0,blend_radius_m)
  movel([0.132597, -1.463646, -2.501823, -0.746921, 1.570796, 1.703394],accel_mss,speed_ms,0,blend_radius_m)
  movel([0.133870, -1.461854, -2.503310, -0.747226, 1.570796, 1.704666],accel_mss,speed_ms,0,blend_radius_m)
  movel([0.135254, -1.460101, -2.504759, -0.747529, 1.570796, 1.706050],accel_mss,speed_ms,0,blend_radius_m)
  movel([0.136763, -1.458395, -2.506165, -0.747828, 1.570796, 1.707560],accel_mss,speed_ms,0,blend_radius_m)
  movel([0.138393, -1.456838, -2.507446, -0.748105, 1.570796, 1.709189],accel_mss,speed_ms,0,blend_radius_m)
  movel([0.143613, -1.452626, -2.510889, -0.748874, 1.570796, 1.714409],accel_mss,speed_ms,0,blend_radius_m)
  movel([0.147757, -1.448828, -2.513971, -0.749590, 1.570796, 1.718554],accel_mss,speed_ms,0,blend_radius_m)
  movel([0.151825, -1.444914, -2.517124, -0.750351, 1.570796, 1.722621],accel_mss,speed_ms,0,blend_radius_m)
  movel([0.153633, -1.443123, -2.518559, -0.750707, 1.570796, 1.724429],accel_mss,speed_ms,0,blend_radius_m)
  speed_ms = 0.005
  movel([0.153633, -1.435007, -2.514811, -0.762571, 1.570796, 1.724429],accel_mss,speed_ms,0,blend_radius_m)
  speed_ms = 0.040
  movel([0.116971, -1.466343, -2.489321, -0.756725, 1.570796, 1.687768],accel_mss,speed_ms,0,blend_radius_m)
  speed_ms = 0.005
  movel([0.116971, -1.474226, -2.492942, -0.745221, 1.570796, 1.687768],accel_mss,speed_ms,0,blend_radius_m)
  speed_ms = 0.025
  movel([0.118906, -1.477174, -2.490437, -0.744779, 1.570796, 1.689702],accel_mss,speed_ms,0,blend_radius_m)
  movel([0.119820, -1.478819, -2.489032, -0.744537, 1.570796, 1.690616],accel_mss,speed_ms,0,blend_radius_m)
  movel([0.120603, -1.480564, -2.487539, -0.744286, 1.570796, 1.691399],accel_mss,speed_ms,0,blend_radius_m)
  movel([0.121192, -1.482390, -2.485971, -0.744028, 1.570796, 1.691988],accel_mss,speed_ms,0,blend_radius_m)
  movel([0.121518, -1.484281, -2.484341, -0.743767, 1.570796, 1.692314],accel_mss,speed_ms,0,blend_radius_m)
  movel([0.121515, -1.486226, -2.482659, -0.743504, 1.570796, 1.692311],accel_mss,speed_ms,0,blend_radius_m)
  movel([0.121368, -1.487215, -2.481802, -0.743372, 1.570796, 1.692164],accel_mss,speed_ms,0,blend_radius_m)
  movel([0.121115, -1.488209, -2.480939, -0.743241, 1.570796, 1.691911],accel_mss,speed_ms,0,blend_radius_m)
  movel([0.120578, -1.487763, -2.481326, -0.743300, 1.570796, 1.691374],accel_mss,speed_ms,0,blend_radius_m)
  movel([0.120282, -1.487237, -2.481783, -0.743369, 1.570796, 1.691079],accel_mss,speed_ms,0,blend_radius_m)
  movel([0.119683, -1.486021, -2.482837, -0.743531, 1.570796, 1.690479],accel_mss,speed_ms,0,blend_radius_m)
  movel([0.118730, -1.484921, -2.483788, -0.743680, 1.570796, 1.689526],accel_mss,speed_ms,0,blend_radius_m)
  movel([0.117627, -1.483937, -2.484638, -0.743814, 1.570796, 1.688423],accel_mss,speed_ms,0,blend_radius_m)
  movel([0.116388, -1.483067, -2.485388, -0.743934, 1.570796, 1.687184],accel_mss,speed_ms,0,blend_radius_m)
  movel([0.115028, -1.482313, -2.486036, -0.744039, 1.570796, 1.685825],accel_mss,speed_ms,0,blend_radius_m)
  movel([0.113563, -1.481676, -2.486584, -0.744129, 1.570796, 1.684359],accel_mss,speed_ms,0,blend_radius_m)
  movel([0.112006, -1.481157, -2.487030, -0.744202, 1.570796, 1.682803],accel_mss,speed_ms,0,blend_radius_m)
  movel([0.110372, -1.480759, -2.487372, -0.744258, 1.570796, 1.681168],accel_mss,speed_ms,0,blend_radius_m)
  movel([0.108677, -1.480478, -2.487612, -0.744298, 1.570796, 1.679474],accel_mss,speed_ms,0,blend_radius_m)
  movel([0.107511, -1.480389, -2.487689, -0.744311, 1.570796, 1.678307],accel_mss,speed_ms,0,blend_radius_m)
  movel([0.106559, -1.480442, -2.487644, -0.744304, 1.570796, 1.677355],accel_mss,speed_ms,0,blend_radius_m)
  movel([0.105807, -1.480621, -2.487490, -0.744278, 1.570796, 1.676604],accel_mss,speed_ms,0,blend_radius_m)
  movel([0.105239, -1.480913, -2.487240, -0.744237, 1.570796, 1.676035],accel_mss,speed_ms,0,blend_radius_m)
  movel([0.104833, -1.481305, -2.486903, -0.744181, 1.570796, 1.675630],accel_mss,speed_ms,0,blend_radius_m)
  movel([0.104576, -1.481784, -2.486491, -0.744113, 1.570796, 1.675372],accel_mss,speed_ms,0,blend_radius_m)
  movel([0.104444, -1.482336, -2.486017, -0.744036, 1.570796, 1.675240],accel_mss,speed_ms,0,blend_radius_m)
  movel([0.104424, -1.482948, -2.485491, -0.743951, 1.570796, 1.675220],accel_mss,speed_ms,0,blend_radius_m)
  movel([0.104640, -1.484298, -2.484326, -0.743764, 1.570796, 1.675436],accel_mss,speed_ms,0,blend_radius_m)
  movel([0.106045, -1.488444, -2.480735, -0.743211, 1.570796, 1.676841],accel_mss,speed_ms,0,blend_radius_m)
  movel([0.104768, -1.487245, -2.481776, -0.743368, 1.570796, 1.675565],accel_mss,speed_ms,0,blend_radius_m)
  movel([0.102297, -1.484784, -2.483907, -0.743698, 1.570796, 1.673094],accel_mss,speed_ms,0,blend_radius_m)
  movel([0.100821, -1.483772, -2.484780, -0.743837, 1.570796, 1.671618],accel_mss,speed_ms,0,blend_radius_m)
  movel([0.098973, -1.482878, -2.485551, -0.743960, 1.570796, 1.669769],accel_mss,speed_ms,0,blend_radius_m)
  movel([0.097026, -1.482082, -2.486235, -0.744071, 1.570796, 1.667823],accel_mss,speed_ms,0,blend_radius_m)
  movel([0.093064, -1.480566, -2.487537, -0.744286, 1.570796, 1.663861],accel_mss,speed_ms,0,blend_radius_m)
  movel([0.091159, -1.479737, -2.488247, -0.744405, 1.570796, 1.661955],accel_mss,speed_ms,0,blend_radius_m)
  movel([0.089380, -1.478789, -2.489058, -0.744542, 1.570796, 1.660176],accel_mss,speed_ms,0,blend_radius_m)
  movel([0.087782, -1.477668, -2.490015, -0.744706, 1.570796, 1.658578],accel_mss,speed_ms,0,blend_radius_m)
  movel([0.086420, -1.476315, -2.491167, -0.744906, 1.570796, 1.657217],accel_mss,speed_ms,0,blend_radius_m)
  movel([0.087205, -1.479872, -2.488131, -0.744385, 1.570796, 1.658001],accel_mss,speed_ms,0,blend_radius_m)
  movel([0.087716, -1.481648, -2.486608, -0.744132, 1.570796, 1.658512],accel_mss,speed_ms,0,blend_radius_m)
  movel([0.088403, -1.483183, -2.485288, -0.743918, 1.570796, 1.659199],accel_mss,speed_ms,0,blend_radius_m)
  movel([0.086999, -1.481912, -2.486381, -0.744095, 1.570796, 1.657796],accel_mss,speed_ms,0,blend_radius_m)
  movel([0.085406, -1.480811, -2.487327, -0.744251, 1.570796, 1.656202],accel_mss,speed_ms,0,blend_radius_m)
  movel([0.082030, -1.478774, -2.489071, -0.744544, 1.570796, 1.652826],accel_mss,speed_ms,0,blend_radius_m)
  movel([0.080988, -1.478003, -2.489729, -0.744656, 1.570796, 1.651784],accel_mss,speed_ms,0,blend_radius_m)
  movel([0.080097, -1.477144, -2.490462, -0.744783, 1.570796, 1.650893],accel_mss,speed_ms,0,blend_radius_m)
  movel([0.078612, -1.475238, -2.492083, -0.745068, 1.570796, 1.649409],accel_mss,speed_ms,0,blend_radius_m)
  movel([0.077247, -1.473232, -2.493783, -0.745374, 1.570796, 1.648043],accel_mss,speed_ms,0,blend_radius_m)
  movel([0.075668, -1.471307, -2.495409, -0.745673, 1.570796, 1.646464],accel_mss,speed_ms,0,blend_radius_m)
  movel([0.075069, -1.470777, -2.495855, -0.745756, 1.570796, 1.645866],accel_mss,speed_ms,0,blend_radius_m)
  movel([0.074358, -1.470358, -2.496208, -0.745823, 1.570796, 1.645154],accel_mss,speed_ms,0,blend_radius_m)
  movel([0.073519, -1.470151, -2.496382, -0.745855, 1.570796, 1.644316],accel_mss,speed_ms,0,blend_radius_m)
  movel([0.073053, -1.470156, -2.496378, -0.745855, 1.570796, 1.643850],accel_mss,speed_ms,0,blend_radius_m)
  movel([0.072551, -1.470254, -2.496296, -0.745839, 1.570796, 1.643347],accel_mss,speed_ms,0,blend_radius_m)
  movel([0.071993, -1.470463, -2.496120, -0.745806, 1.570796, 1.642789],accel_mss,speed_ms,0,blend_radius_m)
  movel([0.071472, -1.470758, -2.495872, -0.745759, 1.570796, 1.642268],accel_mss,speed_ms,0,blend_radius_m)
  movel([0.070527, -1.471547, -2.495206, -0.745635, 1.570796, 1.641324],accel_mss,speed_ms,0,blend_radius_m)
  movel([0.069714, -1.472503, -2.494400, -0.745486, 1.570796, 1.640511],accel_mss,speed_ms,0,blend_radius_m)
  movel([0.069030, -1.473505, -2.493552, -0.745332, 1.570796, 1.639826],accel_mss,speed_ms,0,blend_radius_m)
  movel([0.068855, -1.471775, -2.495015, -0.745600, 1.570796, 1.639652],accel_mss,speed_ms,0,blend_radius_m)
  movel([0.068521, -1.470138, -2.496393, -0.745857, 1.570796, 1.639317],accel_mss,speed_ms,0,blend_radius_m)
  movel([0.067544, -1.467053, -2.498981, -0.746355, 1.570796, 1.638340],accel_mss,speed_ms,0,blend_radius_m)
  movel([0.066452, -1.464030, -2.501503, -0.746856, 1.570796, 1.637249],accel_mss,speed_ms,0,blend_radius_m)
  movel([0.065606, -1.460844, -2.504145, -0.747400, 1.570796, 1.636402],accel_mss,speed_ms,0,blend_radius_m)
  movel([0.065478, -1.459517, -2.505241, -0.747631, 1.570796, 1.636275],accel_mss,speed_ms,0,blend_radius_m)
  movel([0.065543, -1.458089, -2.506418, -0.747882, 1.570796, 1.636339],accel_mss,speed_ms,0,blend_radius_m)
  movel([0.065769, -1.456584, -2.507654, -0.748151, 1.570796, 1.636565],accel_mss,speed_ms,0,blend_radius_m)
  movel([0.066124, -1.455032, -2.508926, -0.748432, 1.570796, 1.636921],accel_mss,speed_ms,0,blend_radius_m)
  movel([0.067117, -1.451878, -2.511498, -0.749013, 1.570796, 1.637914],accel_mss,speed_ms,0,blend_radius_m)
  movel([0.068280, -1.448841, -2.513960, -0.749588, 1.570796, 1.639076],accel_mss,speed_ms,0,blend_radius_m)
  speed_ms = 0.005
  movel([0.068280, -1.440768, -2.510236, -0.761385, 1.570796, 1.639076],accel_mss,speed_ms,0,blend_radius_m)
  speed_ms = 0.040
  # Splitting Linear movement in 2 (instruction 806: MoveL 765)
  movel([0.095656, -1.401848, -2.540190, -0.770351, 1.570796, 1.666452],accel_mss,speed_ms,0,blend_radius_m)
  movel([0.125435, -1.360605, -2.569540, -0.782244, 1.570796, 1.696231],accel_mss,speed_ms,0,blend_radius_m)
  speed_ms = 0.005
  movel([0.125435, -1.369242, -2.573603, -0.769544, 1.570796, 1.696231],accel_mss,speed_ms,0,blend_radius_m)
  speed_ms = 0.025
  movel([0.124073, -1.370110, -2.573002, -0.769277, 1.570796, 1.694869],accel_mss,speed_ms,0,blend_radius_m)
  movel([0.123940, -1.370313, -2.572862, -0.769214, 1.570796, 1.694736],accel_mss,speed_ms,0,blend_radius_m)
  movel([0.123956, -1.370642, -2.572634, -0.769113, 1.570796, 1.694753],accel_mss,speed_ms,0,blend_radius_m)
  movel([0.124394, -1.371658, -2.571928, -0.768803, 1.570796, 1.695190],accel_mss,speed_ms,0,blend_radius_m)
  movel([0.126627, -1.374871, -2.569688, -0.767830, 1.570796, 1.697423],accel_mss,speed_ms,0,blend_radius_m)
  movel([0.130173, -1.379204, -2.566644, -0.766541, 1.570796, 1.700969],accel_mss,speed_ms,0,blend_radius_m)
  movel([0.134442, -1.384114, -2.563162, -0.765113, 1.570796, 1.705239],accel_mss,speed_ms,0,blend_radius_m)
  movel([0.142888, -1.393498, -2.556411, -0.762480, 1.570796, 1.713684],accel_mss,speed_ms,0,blend_radius_m)
  movel([0.147705, -1.398644, -2.552655, -0.761090, 1.570796, 1.718501],accel_mss,speed_ms,0,blend_radius_m)
  movel([0.148198, -1.399036, -2.552367, -0.760986, 1.570796, 1.718995],accel_mss,speed_ms,0,blend_radius_m)
  movel([0.148794, -1.399320, -2.552158, -0.760911, 1.570796, 1.719590],accel_mss,speed_ms,0,blend_radius_m)
  movel([0.149472, -1.399384, -2.552111, -0.760894, 1.570796, 1.720269],accel_mss,speed_ms,0,blend_radius_m)
  movel([0.149839, -1.399303, -2.552171, -0.760915, 1.570796, 1.720636],accel_mss,speed_ms,0,blend_radius_m)
  movel([0.150221, -1.399124, -2.552302, -0.760963, 1.570796, 1.721017],accel_mss,speed_ms,0,blend_radius_m)
  movel([0.150830, -1.398619, -2.552673, -0.761097, 1.570796, 1.721626],accel_mss,speed_ms,0,blend_radius_m)
  movel([0.151323, -1.398008, -2.553121, -0.761260, 1.570796, 1.722120],accel_mss,speed_ms,0,blend_radius_m)
  movel([0.153756, -1.394461, -2.555711, -0.762217, 1.570796, 1.724553],accel_mss,speed_ms,0,blend_radius_m)
  movel([0.155927, -1.390832, -2.558342, -0.763215, 1.570796, 1.726723],accel_mss,speed_ms,0,blend_radius_m)
  movel([0.157841, -1.387144, -2.560996, -0.764249, 1.570796, 1.728637],accel_mss,speed_ms,0,blend_radius_m)
  movel([0.159519, -1.383420, -2.563656, -0.765313, 1.570796, 1.730315],accel_mss,speed_ms,0,blend_radius_m)
  movel([0.160971, -1.379681, -2.566308, -0.766401, 1.570796, 1.731767],accel_mss,speed_ms,0,blend_radius_m)
  movel([0.162213, -1.375948, -2.568934, -0.767507, 1.570796, 1.733010],accel_mss,speed_ms,0,blend_radius_m)
  movel([0.163259, -1.372245, -2.571520, -0.768624, 1.570796, 1.734055],accel_mss,speed_ms,0,blend_radius_m)
  movel([0.164121, -1.368599, -2.574048, -0.769743, 1.570796, 1.734917],accel_mss,speed_ms,0,blend_radius_m)
  movel([0.164401, -1.366960, -2.575177, -0.770251, 1.570796, 1.735197],accel_mss,speed_ms,0,blend_radius_m)
  movel([0.164509, -1.365459, -2.576209, -0.770721, 1.570796, 1.735305],accel_mss,speed_ms,0,blend_radius_m)
  movel([0.164447, -1.364092, -2.577145, -0.771151, 1.570796, 1.735243],accel_mss,speed_ms,0,blend_radius_m)
  movel([0.164225, -1.362858, -2.577989, -0.771542, 1.570796, 1.735021],accel_mss,speed_ms,0,blend_radius_m)
  movel([0.163845, -1.361756, -2.578741, -0.771893, 1.570796, 1.734641],accel_mss,speed_ms,0,blend_radius_m)
  movel([0.163311, -1.360786, -2.579400, -0.772203, 1.570796, 1.734107],accel_mss,speed_ms,0,blend_radius_m)
  movel([0.162632, -1.359940, -2.579975, -0.772474, 1.570796, 1.733429],accel_mss,speed_ms,0,blend_radius_m)
  movel([0.161811, -1.359219, -2.580464, -0.772707, 1.570796, 1.732607],accel_mss,speed_ms,0,blend_radius_m)
  movel([0.160853, -1.358621, -2.580868, -0.772900, 1.570796, 1.731650],accel_mss,speed_ms,0,blend_radius_m)
  movel([0.159766, -1.358144, -2.581191, -0.773054, 1.570796, 1.730562],accel_mss,speed_ms,0,blend_radius_m)
  movel([0.158552, -1.357783, -2.581435, -0.773171, 1.570796, 1.729348],accel_mss,speed_ms,0,blend_radius_m)
  movel([0.157221, -1.357538, -2.581600, -0.773251, 1.570796, 1.728017],accel_mss,speed_ms,0,blend_radius_m)
  movel([0.154223, -1.357383, -2.581705, -0.773301, 1.570796, 1.725019],accel_mss,speed_ms,0,blend_radius_m)
  movel([0.150822, -1.357655, -2.581521, -0.773213, 1.570796, 1.721619],accel_mss,speed_ms,0,blend_radius_m)
  movel([0.147667, -1.358262, -2.581111, -0.773016, 1.570796, 1.718463],accel_mss,speed_ms,0,blend_radius_m)
  movel([0.144482, -1.359204, -2.580473, -0.772711, 1.570796, 1.715278],accel_mss,speed_ms,0,blend_radius_m)
  movel([0.141275, -1.360440, -2.579636, -0.772314, 1.570796, 1.712072],accel_mss,speed_ms,0,blend_radius_m)
  movel([0.138064, -1.361915, -2.578632, -0.771842, 1.570796, 1.708860],accel_mss,speed_ms,0,blend_radius_m)
  movel([0.134865, -1.363581, -2.577495, -0.771313, 1.570796, 1.705661],accel_mss,speed_ms,0,blend_radius_m)
  movel([0.131684, -1.365389, -2.576257, -0.770743, 1.570796, 1.702480],accel_mss,speed_ms,0,blend_radius_m)
  movel([0.125435, -1.369242, -2.573603, -0.769544, 1.570796, 1.696231],accel_mss,speed_ms,0,blend_radius_m)
  movel([0.124073, -1.370110, -2.573002, -0.769277, 1.570796, 1.694869],accel_mss,speed_ms,0,blend_radius_m)
  movel([0.123940, -1.370313, -2.572862, -0.769214, 1.570796, 1.694736],accel_mss,speed_ms,0,blend_radius_m)
  movel([0.123956, -1.370642, -2.572634, -0.769113, 1.570796, 1.694753],accel_mss,speed_ms,0,blend_radius_m)
  movel([0.124094, -1.370965, -2.572410, -0.769014, 1.570796, 1.694890],accel_mss,speed_ms,0,blend_radius_m)
  speed_ms = 0.005
  movel([0.124094, -1.362339, -2.568354, -0.781695, 1.570796, 1.694890],accel_mss,speed_ms,0,blend_radius_m)
  speed_ms = 0.040
  movel([0.119212, -1.343028, -2.581326, -0.788035, 1.570796, 1.690008],accel_mss,speed_ms,0,blend_radius_m)
  speed_ms = 0.005
  movel([0.119212, -1.351778, -2.585466, -0.775145, 1.570796, 1.690008],accel_mss,speed_ms,0,blend_radius_m)
  speed_ms = 0.025
  movel([0.119468, -1.350241, -2.586490, -0.775658, 1.570796, 1.690264],accel_mss,speed_ms,0,blend_radius_m)
  movel([0.119463, -1.348782, -2.587458, -0.776149, 1.570796, 1.690260],accel_mss,speed_ms,0,blend_radius_m)
  movel([0.119197, -1.347436, -2.588349, -0.776603, 1.570796, 1.689993],accel_mss,speed_ms,0,blend_radius_m)
  movel([0.118676, -1.346234, -2.589143, -0.777012, 1.570796, 1.689472],accel_mss,speed_ms,0,blend_radius_m)
  movel([0.116811, -1.343688, -2.590818, -0.777883, 1.570796, 1.687608],accel_mss,speed_ms,0,blend_radius_m)
  movel([0.116404, -1.342879, -2.591348, -0.778162, 1.570796, 1.687201],accel_mss,speed_ms,0,blend_radius_m)
  movel([0.116182, -1.342043, -2.591895, -0.778451, 1.570796, 1.686978],accel_mss,speed_ms,0,blend_radius_m)
  movel([0.116223, -1.341205, -2.592442, -0.778742, 1.570796, 1.687019],accel_mss,speed_ms,0,blend_radius_m)
  movel([0.116610, -1.340382, -2.592979, -0.779028, 1.570796, 1.687406],accel_mss,speed_ms,0,blend_radius_m)
  movel([0.117398, -1.339547, -2.593523, -0.779320, 1.570796, 1.688194],accel_mss,speed_ms,0,blend_radius_m)
  movel([0.118238, -1.339064, -2.593836, -0.779489, 1.570796, 1.689034],accel_mss,speed_ms,0,blend_radius_m)
  movel([0.119101, -1.338875, -2.593959, -0.779555, 1.570796, 1.689897],accel_mss,speed_ms,0,blend_radius_m)
  movel([0.119955, -1.338917, -2.593932, -0.779540, 1.570796, 1.690752],accel_mss,speed_ms,0,blend_radius_m)
  movel([0.121503, -1.339452, -2.593584, -0.779353, 1.570796, 1.692300],accel_mss,speed_ms,0,blend_radius_m)
  movel([0.122639, -1.340183, -2.593109, -0.779098, 1.570796, 1.693435],accel_mss,speed_ms,0,blend_radius_m)
  movel([0.122564, -1.338346, -2.594302, -0.779740, 1.570796, 1.693360],accel_mss,speed_ms,0,blend_radius_m)
  movel([0.122160, -1.336700, -2.595368, -0.780321, 1.570796, 1.692956],accel_mss,speed_ms,0,blend_radius_m)
  movel([0.120761, -1.333731, -2.597282, -0.781376, 1.570796, 1.691558],accel_mss,speed_ms,0,blend_radius_m)
  movel([0.119253, -1.330758, -2.599185, -0.782445, 1.570796, 1.690049],accel_mss,speed_ms,0,blend_radius_m)
  movel([0.118710, -1.329105, -2.600239, -0.783045, 1.570796, 1.689507],accel_mss,speed_ms,0,blend_radius_m)
  movel([0.118451, -1.327251, -2.601416, -0.783721, 1.570796, 1.689248],accel_mss,speed_ms,0,blend_radius_m)
  movel([0.118464, -1.326003, -2.602206, -0.784180, 1.570796, 1.689260],accel_mss,speed_ms,0,blend_radius_m)
  movel([0.118608, -1.324948, -2.602872, -0.784569, 1.570796, 1.689404],accel_mss,speed_ms,0,blend_radius_m)
  movel([0.118867, -1.324077, -2.603421, -0.784891, 1.570796, 1.689664],accel_mss,speed_ms,0,blend_radius_m)
  movel([0.119228, -1.323387, -2.603855, -0.785147, 1.570796, 1.690024],accel_mss,speed_ms,0,blend_radius_m)
  movel([0.119668, -1.322870, -2.604180, -0.785339, 1.570796, 1.690464],accel_mss,speed_ms,0,blend_radius_m)
  movel([0.120176, -1.322516, -2.604402, -0.785471, 1.570796, 1.690972],accel_mss,speed_ms,0,blend_radius_m)
  movel([0.120729, -1.322319, -2.604526, -0.785544, 1.570796, 1.691525],accel_mss,speed_ms,0,blend_radius_m)
  movel([0.121315, -1.322271, -2.604556, -0.785562, 1.570796, 1.692111],accel_mss,speed_ms,0,blend_radius_m)
  movel([0.121915, -1.322365, -2.604497, -0.785527, 1.570796, 1.692711],accel_mss,speed_ms,0,blend_radius_m)
  movel([0.122509, -1.322593, -2.604354, -0.785442, 1.570796, 1.693305],accel_mss,speed_ms,0,blend_radius_m)
  movel([0.123621, -1.323417, -2.603836, -0.785136, 1.570796, 1.694417],accel_mss,speed_ms,0,blend_radius_m)
  movel([0.124517, -1.324675, -2.603044, -0.784669, 1.570796, 1.695313],accel_mss,speed_ms,0,blend_radius_m)
  movel([0.125063, -1.326303, -2.602016, -0.784069, 1.570796, 1.695859],accel_mss,speed_ms,0,blend_radius_m)
  movel([0.125699, -1.324578, -2.603106, -0.784705, 1.570796, 1.696495],accel_mss,speed_ms,0,blend_radius_m)
  movel([0.126097, -1.322975, -2.604114, -0.785300, 1.570796, 1.696893],accel_mss,speed_ms,0,blend_radius_m)
  movel([0.126308, -1.321468, -2.605059, -0.785862, 1.570796, 1.697105],accel_mss,speed_ms,0,blend_radius_m)
  movel([0.126402, -1.317142, -2.607755, -0.787492, 1.570796, 1.697198],accel_mss,speed_ms,0,blend_radius_m)
  movel([0.126577, -1.314067, -2.609656, -0.788666, 1.570796, 1.697374],accel_mss,speed_ms,0,blend_radius_m)
  movel([0.126809, -1.312748, -2.610467, -0.789173, 1.570796, 1.697605],accel_mss,speed_ms,0,blend_radius_m)
  movel([0.127149, -1.311576, -2.611187, -0.789626, 1.570796, 1.697945],accel_mss,speed_ms,0,blend_radius_m)
  movel([0.127576, -1.310557, -2.611810, -0.790021, 1.570796, 1.698372],accel_mss,speed_ms,0,blend_radius_m)
  movel([0.128074, -1.309694, -2.612338, -0.790357, 1.570796, 1.698870],accel_mss,speed_ms,0,blend_radius_m)
  movel([0.128623, -1.308990, -2.612767, -0.790632, 1.570796, 1.699419],accel_mss,speed_ms,0,blend_radius_m)
  movel([0.129206, -1.308447, -2.613098, -0.790844, 1.570796, 1.700002],accel_mss,speed_ms,0,blend_radius_m)
  movel([0.129804, -1.308069, -2.613329, -0.790992, 1.570796, 1.700600],accel_mss,speed_ms,0,blend_radius_m)
  movel([0.130399, -1.307859, -2.613456, -0.791074, 1.570796, 1.701195],accel_mss,speed_ms,0,blend_radius_m)
  movel([0.130971, -1.307820, -2.613480, -0.791089, 1.570796, 1.701767],accel_mss,speed_ms,0,blend_radius_m)
  movel([0.131502, -1.307955, -2.613398, -0.791037, 1.570796, 1.702299],accel_mss,speed_ms,0,blend_radius_m)
  movel([0.131976, -1.308264, -2.613210, -0.790916, 1.570796, 1.702773],accel_mss,speed_ms,0,blend_radius_m)
  movel([0.132374, -1.308752, -2.612912, -0.790724, 1.570796, 1.703171],accel_mss,speed_ms,0,blend_radius_m)
  movel([0.132675, -1.309422, -2.612504, -0.790463, 1.570796, 1.703472],accel_mss,speed_ms,0,blend_radius_m)
  movel([0.132863, -1.310274, -2.611984, -0.790131, 1.570796, 1.703660],accel_mss,speed_ms,0,blend_radius_m)
  movel([0.132920, -1.311311, -2.611349, -0.789729, 1.570796, 1.703717],accel_mss,speed_ms,0,blend_radius_m)
  movel([0.132831, -1.312531, -2.610601, -0.789257, 1.570796, 1.703628],accel_mss,speed_ms,0,blend_radius_m)
  movel([0.133993, -1.311099, -2.611479, -0.789811, 1.570796, 1.704789],accel_mss,speed_ms,0,blend_radius_m)
  movel([0.134992, -1.309633, -2.612375, -0.790381, 1.570796, 1.705788],accel_mss,speed_ms,0,blend_radius_m)
  movel([0.135861, -1.308138, -2.613286, -0.790965, 1.570796, 1.706657],accel_mss,speed_ms,0,blend_radius_m)
  movel([0.136634, -1.306621, -2.614208, -0.791560, 1.570796, 1.707431],accel_mss,speed_ms,0,blend_radius_m)
  movel([0.139470, -1.300489, -2.617902, -0.793998, 1.570796, 1.710266],accel_mss,speed_ms,0,blend_radius_m)
  movel([0.140575, -1.298227, -2.619253, -0.794909, 1.570796, 1.711371],accel_mss,speed_ms,0,blend_radius_m)
  movel([0.142098, -1.295575, -2.620828, -0.795986, 1.570796, 1.712895],accel_mss,speed_ms,0,blend_radius_m)
  movel([0.143032, -1.294355, -2.621550, -0.796485, 1.570796, 1.713828],accel_mss,speed_ms,0,blend_radius_m)
  movel([0.144085, -1.293342, -2.622147, -0.796900, 1.570796, 1.714882],accel_mss,speed_ms,0,blend_radius_m)
  movel([0.144662, -1.292947, -2.622380, -0.797062, 1.570796, 1.715458],accel_mss,speed_ms,0,blend_radius_m)
  movel([0.145910, -1.292435, -2.622681, -0.797273, 1.570796, 1.716706],accel_mss,speed_ms,0,blend_radius_m)
  movel([0.146584, -1.292350, -2.622731, -0.797308, 1.570796, 1.717380],accel_mss,speed_ms,0,blend_radius_m)
